// TIA Portal project "UsineEcole_TIAV20" (V20)

(* hardware
DEVICE "Station S71500/ET200MP_1"  S7-1500 station
   slot 0: "Châssis_0"  Rack  6ES7 590-1***0-0AA0
   slot 1: "PLC_1"  CPU 1518-4 PN/DP  6ES7 518-4AP00-0AB0  V2.9
      slot 3: "Ecran CPU_1"  6ES7591-1BA00-0AA0
      slot 32768: "Interface PROFINET_1"  X1
      slot 33024: "Interface PROFINET_2"  X2
      slot 33280: "Interface PROFINET GBIT_3"  X3
      slot 34817: "Virtual CP interface port_1"  Virtual CP interface port  Virtual CP interface port
   slot 2: "DI 32x24VDC HF_1"  DI 32x24VDC HF  6ES7 521-1BL00-0AB0  V2.1
   slot 3: "DQ 32x24VDC/0.5A ST_1"  DQ 32x24VDC/0.5A ST  6ES7 522-1BL00-0AB0  V2.0
DEVICE "Appareil GSD_1"  GSD.Device.PN
   slot 0: "Châssis"  Rack  V1.0
   slot 0: "REP 1"  AL1306  AL1306
      slot 0: "PROFINET interface"  PROFINET interface
      slot 1: "PN-IO"  PN-IO
         slot 1: "X21"  X21
         slot 2: "X22"  X22
   slot 1: "IO-Link  1 I Byte without PQI"  IO-Link  1 I Byte without PQI
   slot 1: "Digital Input"  Digital Input
   slot 1: "8 Ports - IO Mode_1"  8 Ports - IO Mode
      slot 0: "IO-Link Master Proxy"  IO-Link Master Proxy
   slot 1: "Digital Input without PD"  Digital Input without PD
   slot 2: "IO-Link  1 I Byte without PQI_1"  IO-Link  1 I Byte without PQI
   slot 2: "Digital Input_1"  Digital Input
   slot 2: "Digital Input without PD_1"  Digital Input without PD
   slot 3: "IO-Link  1 I Byte without PQI_2"  IO-Link  1 I Byte without PQI
   slot 3: "Digital Input_2"  Digital Input
   slot 3: "Digital Input without PD_2"  Digital Input without PD
   slot 4: "IO-Link  1 I Byte without PQI_3"  IO-Link  1 I Byte without PQI
   slot 4: "Digital Input_3"  Digital Input
   slot 4: "Digital Input without PD_3"  Digital Input without PD
   slot 5: "IO-Link  1 I Byte without PQI_4"  IO-Link  1 I Byte without PQI
   slot 5: "Digital Input_4"  Digital Input
   slot 5: "Digital Input without PD_4"  Digital Input without PD
   slot 6: "IO-Link  1 I Byte without PQI_5"  IO-Link  1 I Byte without PQI
   slot 6: "Digital Input_5"  Digital Input
   slot 6: "Digital Input without PD_5"  Digital Input without PD
   slot 7: "IO-Link  1 I Byte without PQI_6"  IO-Link  1 I Byte without PQI
   slot 7: "Digital Input_6"  Digital Input
   slot 7: "Digital Input without PD_6"  Digital Input without PD
   slot 8: "IO-Link  1 I Byte without PQI_7"  IO-Link  1 I Byte without PQI
   slot 8: "Digital Input_7"  Digital Input
   slot 8: "Digital Input without PD_7"  Digital Input without PD
DEVICE "Appareil GSD_2"  GSD.Device.PN
   slot 0: "Châssis"  Rack  V1.0
   slot 0: "REP 2"  AL1306  AL1306
      slot 0: "PROFINET interface"  PROFINET interface
      slot 1: "PN-IO"  PN-IO
         slot 1: "X21"  X21
         slot 2: "X22"  X22
   slot 1: "8 Ports - IO Mode_1"  8 Ports - IO Mode
      slot 0: "IO-Link Master Proxy"  IO-Link Master Proxy
   slot 1: "Digital Input without PD"  Digital Input without PD
   slot 2: "Digital Input without PD_1"  Digital Input without PD
   slot 3: "Digital Input without PD_2"  Digital Input without PD
   slot 4: "Digital Input without PD_3"  Digital Input without PD
   slot 5: "Digital Input without PD_4"  Digital Input without PD
   slot 6: "Digital Input without PD_5"  Digital Input without PD
   slot 7: "Digital Input without PD_6"  Digital Input without PD
   slot 8: "Digital Input without PD_7"  Digital Input without PD
DEVICE "Appareil GSD_3"  GSD.Device.PN
   slot 0: "Châssis"  Rack  V1.0
   slot 0: "REP 3"  AL1306  AL1306
      slot 0: "PROFINET interface"  PROFINET interface
      slot 1: "PN-IO"  PN-IO
         slot 1: "X21"  X21
         slot 2: "X22"  X22
   slot 1: "8 Ports - IO Mode_1"  8 Ports - IO Mode
      slot 0: "IO-Link Master Proxy"  IO-Link Master Proxy
   slot 1: "Digital Input without PD"  Digital Input without PD
   slot 2: "Digital Input without PD_1"  Digital Input without PD
   slot 3: "Digital Input without PD_2"  Digital Input without PD
   slot 4: "Digital Input without PD_3"  Digital Input without PD
   slot 5: "Digital Input without PD_4"  Digital Input without PD
   slot 6: "Digital Input without PD_5"  Digital Input without PD
   slot 7: "Digital Input without PD_6"  Digital Input without PD
   slot 8: "Digital Input without PD_7"  Digital Input without PD
DEVICE "Appareil GSD_4"  GSD.Device.PN
   slot 0: "Châssis"  Rack  V1.0
   slot 0: "REP 4"  AL1306  AL1306
      slot 0: "PROFINET interface"  PROFINET interface
      slot 1: "PN-IO"  PN-IO
         slot 1: "X21"  X21
         slot 2: "X22"  X22
   slot 1: "8 Ports - IO Mode_1"  8 Ports - IO Mode
      slot 0: "IO-Link Master Proxy"  IO-Link Master Proxy
   slot 1: "Digital Input without PD"  Digital Input without PD
   slot 2: "Digital Input without PD_1"  Digital Input without PD
   slot 3: "Digital Input without PD_2"  Digital Input without PD
   slot 4: "Digital Input without PD_3"  Digital Input without PD
   slot 5: "Digital Input without PD_4"  Digital Input without PD
   slot 6: "Digital Input without PD_5"  Digital Input without PD
   slot 7: "Digital Input without PD_6"  Digital Input without PD
   slot 8: "Digital Input without PD_7"  Digital Input without PD
DEVICE "Appareil GSD_5"  GSD.Device.PN
   slot 0: "Châssis"  Rack  V1.0
   slot 0: "REP 5"  AL1306  AL1306
      slot 0: "PROFINET interface"  PROFINET interface
      slot 1: "PN-IO"  PN-IO
         slot 1: "X21"  X21
         slot 2: "X22"  X22
   slot 1: "8 Ports - IO Mode_1"  8 Ports - IO Mode
      slot 0: "IO-Link Master Proxy"  IO-Link Master Proxy
   slot 1: "Digital Input without PD"  Digital Input without PD
   slot 2: "Digital Input without PD_1"  Digital Input without PD
   slot 3: "Digital Input without PD_2"  Digital Input without PD
   slot 4: "Digital Input without PD_3"  Digital Input without PD
   slot 5: "Digital Input without PD_4"  Digital Input without PD
   slot 6: "Digital Input without PD_5"  Digital Input without PD
   slot 7: "Digital Input without PD_6"  Digital Input without PD
   slot 8: "Digital Input without PD_7"  Digital Input without PD
DEVICE "Appareil GSD_6"  GSD.Device.PN
   slot 0: "Châssis"  Rack  V1.0
   slot 0: "REP 6"  AL1306  AL1306
      slot 0: "PROFINET interface"  PROFINET interface
      slot 1: "PN-IO"  PN-IO
         slot 1: "X21"  X21
         slot 2: "X22"  X22
   slot 1: "8 Ports - IO Mode_1"  8 Ports - IO Mode
      slot 0: "IO-Link Master Proxy"  IO-Link Master Proxy
   slot 1: "Digital Input without PD"  Digital Input without PD
   slot 2: "Digital Input without PD_1"  Digital Input without PD
   slot 3: "Digital Input without PD_2"  Digital Input without PD
   slot 4: "Digital Input without PD_3"  Digital Input without PD
   slot 5: "Digital Input without PD_4"  Digital Input without PD
   slot 6: "Digital Input without PD_5"  Digital Input without PD
   slot 7: "Digital Input without PD_6"  Digital Input without PD
   slot 8: "Digital Input without PD_7"  Digital Input without PD
DEVICE "Appareil GSD_7"  GSD.Device.PN
   slot 0: "Châssis"  Rack  V1.0
   slot 0: "Ilot 01"  EX260 SPN 1/2  EX260-SPN
      slot 0: "EX260 SPN 1/2"  EX260 SPN 1/2
      slot 1: "Interface"  Interface
         slot 1: "Port 1 - RJ45"  Port 1 - RJ45
         slot 2: "Port 2 - RJ45"  Port 2 - RJ45
      slot 1: "  4 byte  Output_1"    4 byte  Output
         slot 0: "  4 byte  Output"    4 byte  Output
DEVICE "Appareil GSD_8"  GSD.Device.PN
   slot 0: "Châssis"  Rack  V1.0
   slot 0: "ilot02"  EX260 SPN 1/2  EX260-SPN
      slot 0: "EX260 SPN 1/2"  EX260 SPN 1/2
      slot 1: "Interface"  Interface
         slot 1: "Port 1 - RJ45"  Port 1 - RJ45
         slot 2: "Port 2 - RJ45"  Port 2 - RJ45
      slot 1: "  4 byte  Output_1"    4 byte  Output
         slot 0: "  4 byte  Output"    4 byte  Output
DEVICE "Appareil GSD_9"  GSD.Device.PN
   slot 0: "Châssis"  Rack  V1.0
   slot 0: "SP-COP2-ENI"  R1.190.1320.0  R1.190.1320.0
      slot 0: "R1.190.1320.0"  R1.190.1320.0
      slot 1: "SP-COP2-ENI Diagnostics"  SP-COP2-ENI Diagnostics
      slot 2: "jz"  Interface
         slot 1: "RJ45 10/100 MBit/s"  RJ45 10/100 MBit/s
   slot 16: "Logic input block 1_1"  Logic input block 1
      slot 0: "Logic input block 1"  Logic input block 1
   slot 21: "Logic output block 1_1"  Logic output block 1
      slot 0: "Logic output block 1"  Logic output block 1
   slot 32: "CRC data_1"  CRC data
      slot 0: "CRC data"  CRC data
   slot 33: "Status data_1"  Status data
      slot 0: "Status data"  Status data
   slot 34: "Auxiliary data_1"  Auxiliary data
      slot 0: "Auxiliary data"  Auxiliary data
DEVICE "HMI_1"  TP1500 Comfort
   slot 0: "HMI_1"  TP1500 Comfort  6AV2 124-0QC02-0AX1  17.0.0.0
   slot 1: "HMI_RT_1"  TP1500 Comfort  6AV2 124-0QC02-0AX1  17.0.0.0
   slot 5: "HMI_1.IE_CP_1"  PROFINET Interface  17.0.0.0
      slot 1: "Interface PROFINET_1"  PROFINET Interface
         slot 1: "Port_1"  Port
         slot 2: "Port_2"  Port
   slot 6: "HMI_1.IE_CP_2"  PROFINET Interface  17.0.0.0
      slot 1: "Interface PROFINET_GBit"  PROFINET Interface
         slot 1: "Port_1"  Port
   slot 7: "HMI_1.MPI/DP_CP_1"  MPI/DP Interface  17.0.0.0
DEVICE "SINAMICS G_1"  Sinamics.Device
   slot 0: "	_0"  Rail  SinamicsG120CRackP
   slot 0: "Convoyeur 01"  G120C PN  6SL3210-1KE11-8UF2  4.7.13
      slot 1: "Interface PROFINET"  MDD-SinamicsG120-P
      slot 3: "PM G120C"  PM G120C  6SL3210-1KE11-8UF2  -
DEVICE "SINAMICS G_2"  Sinamics.Device
   slot 0: "	_0"  Rail  SinamicsG120CRackP
   slot 0: "Convoyeur 02"  G120C PN  6SL3210-1KE11-8UF2  4.7.13
      slot 1: "Interface PROFINET"  MDD-SinamicsG120-P
      slot 3: "PM G120C"  PM G120C  6SL3210-1KE11-8UF2  -
DEVICE "SINAMICS G_3"  Sinamics.Device
   slot 0: "	_0"  Rail  SinamicsG120CRackP
   slot 0: "Convoyeur 03"  G120C PN  6SL3210-1KE11-8UF2  4.7.13
      slot 1: "Interface PROFINET"  MDD-SinamicsG120-P
      slot 3: "PM G120C"  PM G120C  6SL3210-1KE11-8UF2  -
DEVICE "Appareil GSD_10"  GSD.Device
   slot 0: "Châssis_0"  Rail
DEVICE "Appareil GSD_12"  GSD.Device.PN
   slot 0: "Châssis"  Rack  V1.0
   slot 0: "UR_R4"  V1.0  0000201
      slot 0: "V1.0"  V1.0
      slot 1: "Interface"  Interface
         slot 1: "RJ45 10/100 MBit/s"  RJ45 10/100 MBit/s
   slot 1: "1_T2O State_1"  1_T2O State  1.0
      slot 0: "1_T2O State"  1_T2O State
   slot 2: "2_T2O IO_1"  2_T2O IO  1.0
      slot 0: "2_T2O IO"  2_T2O IO
   slot 3: "3_T2O Joints_1"  3_T2O Joints  1.0
      slot 0: "3_T2O Joints"  3_T2O Joints
   slot 4: "4_T2O TCP_1"  4_T2O TCP  1.0
      slot 0: "4_T2O TCP"  4_T2O TCP
   slot 5: "5_T2O General Purpose Bit Registers_1"  5_T2O General Purpose Bit Registers  1.0
      slot 0: "5_T2O General Purpose Bit Registers"  5_T2O General Purpose Bit Registers
   slot 6: "6_T2O General Purpose Int Registers_1"  6_T2O General Purpose Int Registers  1.0
      slot 0: "6_T2O General Purpose Int Registers"  6_T2O General Purpose Int Registers
   slot 7: "7_T2O General Purpose Float Registers_1"  7_T2O General Purpose Float Registers  1.0
      slot 0: "7_T2O General Purpose Float Registers"  7_T2O General Purpose Float Registers
   slot 8: "8_O2T Robot IO_1"  8_O2T Robot IO  1.0
      slot 0: "8_O2T Robot IO"  8_O2T Robot IO
   slot 9: "9_O2T General Purpose Registers 1_1"  9_O2T General Purpose Registers 1  1.0
      slot 0: "9_O2T General Purpose Registers 1"  9_O2T General Purpose Registers 1
   slot 10: "10_O2T General Purpose Registers 2_1"  10_O2T General Purpose Registers 2  1.0
      slot 0: "10_O2T General Purpose Registers 2"  10_O2T General Purpose Registers 2
DEVICE "Appareil GSD_13"  GSD.Device.PN
   slot 0: "Châssis"  Rack  V1.0
   slot 0: "URIODev1_1"  V1.0  0000201
      slot 0: "V1.0"  V1.0
      slot 1: "Interface"  Interface
         slot 1: "RJ45 10/100 MBit/s"  RJ45 10/100 MBit/s
   slot 1: "1_T2O State_1"  1_T2O State  1.0
      slot 0: "1_T2O State"  1_T2O State
   slot 2: "2_T2O IO_1"  2_T2O IO  1.0
      slot 0: "2_T2O IO"  2_T2O IO
   slot 3: "3_T2O Joints_1"  3_T2O Joints  1.0
      slot 0: "3_T2O Joints"  3_T2O Joints
   slot 4: "4_T2O TCP_1"  4_T2O TCP  1.0
      slot 0: "4_T2O TCP"  4_T2O TCP
   slot 5: "5_T2O General Purpose Bit Registers_1"  5_T2O General Purpose Bit Registers  1.0
      slot 0: "5_T2O General Purpose Bit Registers"  5_T2O General Purpose Bit Registers
   slot 6: "6_T2O General Purpose Int Registers_1"  6_T2O General Purpose Int Registers  1.0
      slot 0: "6_T2O General Purpose Int Registers"  6_T2O General Purpose Int Registers
   slot 7: "7_T2O General Purpose Float Registers_1"  7_T2O General Purpose Float Registers  1.0
      slot 0: "7_T2O General Purpose Float Registers"  7_T2O General Purpose Float Registers
   slot 8: "8_O2T Robot IO_1"  8_O2T Robot IO  1.0
      slot 0: "8_O2T Robot IO"  8_O2T Robot IO
   slot 9: "9_O2T General Purpose Registers 1_1"  9_O2T General Purpose Registers 1  1.0
      slot 0: "9_O2T General Purpose Registers 1"  9_O2T General Purpose Registers 1
   slot 10: "10_O2T General Purpose Registers 2_1"  10_O2T General Purpose Registers 2  1.0
      slot 0: "10_O2T General Purpose Registers 2"  10_O2T General Purpose Registers 2
   slot 11: "PROFIsafe_1"  PROFIsafe  1.0
      slot 0: "Module Access Point"  Module Access Point
DEVICE "Appareil GSD_11"  GSD.Device.PN
   slot 0: "Châssis"  Rack  V1.0
   slot 0: "CP-1604"  V2.5  A05B-2500-J930  V2.5
      slot 0: "CP 1604"  CP 1604
      slot 1: "Interface"  Interface
         slot 1: "Port_1"  Port
   slot 1: "  32 octets_1"  32 bytes  1.0
      slot 0: "  32 octets"  32 bytes
DEVICE "Appareil GSD_14"  GSD.Device.PN
   slot 0: "Châssis"  Rack  V1.0
   slot 0: "cv-x400"  CV-X4XX  CV-X4XX  5.1
      slot 0: "CV-X4XX"  CV-X4XX  5.1
      slot 1: "Interface"  Interface
         slot 1: "Port 1"  Port 1
   slot 1: "Command and Result Status_1"  Command and Result Status
      slot 0: "Command and Result Status"  Command and Result Status
   slot 2: "Trg Ready Status_1"  Trg Ready Status
      slot 0: "Trg Ready Status"  Trg Ready Status
   slot 3: "Trg Ack Status_1"  Trg Ack Status
      slot 0: "Trg Ack Status"  Trg Ack Status
   slot 4: "Miscellaneous Status_1"  Miscellaneous Status
      slot 0: "Miscellaneous Status"  Miscellaneous Status
   slot 5: "Tool Judge Value_1"  Tool Judge Value
      slot 0: "Tool Judge Value"  Tool Judge Value
   slot 6: "Result Data 128Byte_1"  Result Data 128Byte
      slot 0: "Result Data 128Byte"  Result Data 128Byte
   slot 7: "Result Data 32Byte_1"  Result Data 32Byte
      slot 0: "Result Data 32Byte"  Result Data 32Byte
   slot 8: "Result Data 32Byte_2"  Result Data 32Byte
      slot 0: "Result Data 32Byte"  Result Data 32Byte
   slot 9: "Result Data 32Byte_3"  Result Data 32Byte
      slot 0: "Result Data 32Byte"  Result Data 32Byte
   slot 10: "Result Data 32Byte_4"  Result Data 32Byte
      slot 0: "Result Data 32Byte"  Result Data 32Byte
   slot 11: "Result Data 32Byte_5"  Result Data 32Byte
      slot 0: "Result Data 32Byte"  Result Data 32Byte
   slot 12: "Command and Result Control_1"  Command and Result Control
      slot 0: "Command and Result Control"  Command and Result Control
   slot 13: "Trg Control_1"  Trg Control
      slot 0: "Trg Control"  Trg Control
   slot 14: "Miscellaneous Control_1"  Miscellaneous Control
      slot 0: "Miscellaneous Control"  Miscellaneous Control
   slot 15: "Reserved Control_1"  Reserved Control
      slot 0: "Reserved Control"  Reserved Control
   slot 16: "Reserved Control_2"  Reserved Control
      slot 0: "Reserved Control"  Reserved Control
   slot 17: "Parameter 128Byte_1"  Parameter 128Byte
      slot 0: "Parameter 128Byte"  Parameter 128Byte
   slot 18: "Parameter 32Byte_1"  Parameter 32Byte
      slot 0: "Parameter 32Byte"  Parameter 32Byte
   slot 19: "Parameter 32Byte_2"  Parameter 32Byte
      slot 0: "Parameter 32Byte"  Parameter 32Byte
   slot 20: "Parameter 32Byte_3"  Parameter 32Byte
      slot 0: "Parameter 32Byte"  Parameter 32Byte
   slot 21: "Parameter 32Byte_4"  Parameter 32Byte
      slot 0: "Parameter 32Byte"  Parameter 32Byte
   slot 22: "Parameter 32Byte_5"  Parameter 32Byte
      slot 0: "Parameter 32Byte"  Parameter 32Byte
DEVICE "GSD device_1"  GSD.Device.PN
   slot 0: "Rack"  Rack  V1.0
   slot 0: "REP 4_rep"  AL1102  AL1102
      slot 0: "AL1102"  AL1102
      slot 1: "X1"  X1
         slot 1: "Port 1"  Port 1
         slot 2: "Port 2"  Port 2
      slot 1: "8 Ports_1"  8 Ports  AL1102
         slot 0: "IO-Link Master"  IO-Link Master
   slot 1: "Digital Input + PQI"  Digital Input + PQI
   slot 2: "Digital Input + PQI_1"  Digital Input + PQI
DEVICE "GSD device_2"  GSD.Device.PN
   slot 0: "Rack"  Rack  V1.0
   slot 0: "OmniCore"  OmniCore Standard  3020-x  V1.1
      slot 0: "OmniCore Standard PROFINET Device"  OmniCore Standard PROFINET Device
      slot 1: "PROFINET Interface"  PROFINET Interface
         slot 1: "Network Port 1"  Network Port 1
   slot 1: "DI 8 bytes_1"  DI 8 bytes
      slot 0: "DI 8 bytes"  DI 8 bytes
   slot 2: "DO 8 bytes_1"  DO 8 bytes
      slot 0: "DO 8 bytes"  DO 8 bytes
*)

// ===== PLC "PLC_1"  CPU 1518-4 PN/DP =====

VAR_GLOBAL   // PLC tag table "Table de variables standard"
   "I_En_Service" AT %I0.0 : Bool;
   "I_Not_AU" AT %I0.1 : Bool;   // Entree AU: 1 = pas d'arret d'urgence
   "I_En_Manuel" AT %I0.2 : Bool;
   "I_En_Automatique" AT %I0.3 : Bool;
   "I_porte_non_réarmée" AT %I0.4 : Bool;
   "I_porte_01_Op" AT %I0.5 : Bool;
   "I_porte_02_Op" AT %I0.6 : Bool;
   "I_libre_I07" AT %I0.7 : Bool;
   "I_libre_I10" AT %I1.0 : Bool;
   "I_Def_Thermique_CV01_hyppo" AT %I1.1 : Bool;
   "I_Def_Thermique_CV02_hyppo" AT %I1.2 : Bool;
   "I_Def_Thermique_CV03_hyppo" AT %I1.3 : Bool;
   "I_Def_Thermique_CV04_hyppo" AT %I1.4 : Bool;
   "I_libre_I15" AT %I1.5 : Bool;
   "I_libre_I16" AT %I1.6 : Bool;
   "I_libre_I17" AT %I1.7 : Bool;
   "I_libre_I20" AT %I2.0 : Bool;
   "I_libre_I21" AT %I2.1 : Bool;
   "I_libre_I22" AT %I2.2 : Bool;
   "I_libre_I23" AT %I2.3 : Bool;
   "I_libre_I24" AT %I2.4 : Bool;
   "I_libre_I25" AT %I2.5 : Bool;
   "I_libre_I26" AT %I2.6 : Bool;
   "I_libre_I27" AT %I2.7 : Bool;
   "I_libre_I30" AT %I3.0 : Bool;
   "I_libre_I31" AT %I3.1 : Bool;
   "I_libre_I32" AT %I3.2 : Bool;
   "I_libre_I33" AT %I3.3 : Bool;
   "I_libre_I34" AT %I3.4 : Bool;
   "I_libre_I35" AT %I3.5 : Bool;
   "I_libre_I36" AT %I3.6 : Bool;
   "I_libre_I37" AT %I3.7 : Bool;
   "I_Pres_Pal_B01" AT %I5.0 : Bool;
   "I_Pres_Elev_B01" AT %I4.0 : Bool;
   "I_Elev_01_Bas" AT %I5.1 : Bool;
   "I_Elev_01_Haut" AT %I4.1 : Bool;
   "I_Pres_Pal_B02" AT %I5.2 : Bool;
   "I_Pres_Elev_B02" AT %I4.2 : Bool;
   "I_Elev_02_Bas" AT %I5.3 : Bool;
   "I_Elev_02_Haut" AT %I4.3 : Bool;
   "I_Pres_Pal_B03" AT %I5.4 : Bool;
   "I_Pres_Elev_B03" AT %I4.4 : Bool;
   "I_Elev_03_Bas" AT %I5.5 : Bool;
   "I_Elev_03_Haut" AT %I4.5 : Bool;
   "I_Pres_Pal_B04" AT %I5.6 : Bool;
   "I_Pres_Elev_B04" AT %I4.6 : Bool;
   "I_Elev_04_Bas" AT %I5.7 : Bool;
   "I_Elev_04_Haut" AT %I4.7 : Bool;
   "I_Pres_Pal_B05" AT %I7.0 : Bool;
   "I_Pres_Elev_B05" AT %I6.0 : Bool;
   "I_Elev_05_Bas" AT %I7.1 : Bool;
   "I_Elev_05_Haut" AT %I6.1 : Bool;
   "I_Pres_Pal_B06" AT %I7.2 : Bool;
   "I_Pres_Elev_B06" AT %I6.2 : Bool;
   "I_Elev_06_Bas" AT %I7.3 : Bool;
   "I_Elev_06_Haut" AT %I6.3 : Bool;
   "I_Pres_Pal_B07" AT %I7.4 : Bool;
   "I_Pres_Elev_B07" AT %I6.4 : Bool;
   "I_Elev_07_Bas" AT %I7.5 : Bool;
   "I_Elev_07_Haut" AT %I6.5 : Bool;
   "I_det_Phot_01" AT %I11.0 : Bool;
   "I_det_Phot_02" AT %I10.0 : Bool;
   "I_det_Phot_03" AT %I11.1 : Bool;
   "I_verin_blocage_boite_sorti_01" AT %I10.1 : Bool;
   "I_verin_blocage_boite_rentré_01" AT %I11.2 : Bool;
   "I_verin_blocage_boite_sorti_02" AT %I10.2 : Bool;
   "I_verin_blocage_boite_sorti_03" AT %I10.3 : Bool;
   "I_verin_blocage_boite_rentré_03" AT %I11.4 : Bool;
   "I_verin_blocage_boite_rentré_02" AT %I11.3 : Bool;
   "I_verin_blocage_boite_sorti_04" AT %I10.4 : Bool;
   "I_verin_blocage_boite_rentré_04" AT %I11.5 : Bool;
   "I_Det_Phot_04" AT %I13.0 : Bool;
   "I_Det_Phot_05" AT %I12.0 : Bool;
   "I_Det_Phot_06" AT %I13.1 : Bool;
   "I_Det_Photo_7" AT %I15.0 : Bool;
   "I_Det_Photo_8" AT %I14.0 : Bool;
   "I_Det_Photo_9" AT %I15.1 : Bool;
   "I_Wieland_Au_armoire" AT %I16.0 : Bool;
   "I_Wieland_Au_porte01" AT %I16.1 : Bool;
   "I_Wieland_Au_Porte02" AT %I16.2 : Bool;
   "I_Wieland_Au_Robot01_Fanuc" AT %I16.3 : Bool;
   "I_Wieland_Au_Robot02_Fanuc" AT %I16.4 : Bool;
   "I_Wieland_Au_Robot03_ABB" AT %I16.5 : Bool;
   "I_Wielmand_Au_Robot04_UR" AT %I16.6 : Bool;
   "I_Wieland_Au_Robot05_UR" AT %I16.7 : Bool;
   "I_wieland_Au_Carroussel" AT %I17.0 : Bool;
   "I_Wieland_Au_Carterisation" AT %I17.1 : Bool;
   "I_Wieland_Porte 01 ouverte" AT %I17.2 : Bool;
   "I_Wieland_Porte 02 Ouverte" AT %I17.3 : Bool;
   "I_Wieland_Rearmement" AT %I17.4 : Bool;
   "I_Wieland_Dmd acces" AT %I17.5 : Bool;
   "I_Wieland_Mise sous puissance" AT %I17.6 : Bool;
   "I_Wieland_Mise hors puissance" AT %I17.7 : Bool;
   "I_Wieland_Acces_autorisé" AT %I18.0 : Bool;
   "I_Wieland_rearmement_Porte" AT %I18.1 : Bool;
   "I_Wieland_En_Service" AT %I18.2 : Bool;
   "I_Wieland_Porte_non_Réarmée" AT %I18.3 : Bool;
   "I_porte_vision_op" AT %I7.6 : Bool;
   "I_porte_vision_cl" AT %I6.6 : Bool;
   "Tag_1" AT %I590.0 : Bool;
   "Tag_2" AT %I590.1 : Bool;
   "UR01I" AT %I556.0 : "UR__T2O_IOs";
   "Fanuc01_Selecteur_Auto" AT %I30.4 : Bool;
   "Fanuc02_Selecteur_Auto" AT %I220.4 : Bool;
   "Fanuc02_reception_signal_pret" AT %I30.5 : Bool;
   "Fanuc01_reception_signal_pret" AT %I220.5 : Bool;
   "VisionOK" AT %I42.0 : Bool;   // vision OK
   "Tag_8" AT %I42.1 : Bool;
   "Tag_9" AT %I42.2 : Bool;
   "Tag_10" AT %I7.7 : Bool;
   "O_CL_verte" AT %Q0.0 : Bool;
   "O_CL_Orange" AT %Q0.1 : Bool;
   "O_CL_Rouge" AT %Q0.2 : Bool;
   "Q_LibreQ03" AT %Q0.3 : Bool;
   "Q_LibreQ04" AT %Q0.4 : Bool;
   "Q_LibreQ05" AT %Q0.5 : Bool;
   "Q_LibreQ06" AT %Q0.6 : Bool;
   "Q_LibreQ07" AT %Q0.7 : Bool;
   "Q_LibreQ10" AT %Q1.0 : Bool;
   "Q_LibreQ11" AT %Q1.1 : Bool;
   "Q_LibreQ12" AT %Q1.2 : Bool;
   "Q_LibreQ13" AT %Q1.3 : Bool;
   "Q_LibreQ14" AT %Q1.4 : Bool;
   "Q_LibreQ15" AT %Q1.5 : Bool;
   "Q_LibreQ16" AT %Q1.6 : Bool;
   "Q_LibreQ17" AT %Q1.7 : Bool;
   "O_ON_CV_01_Hyppo" AT %Q2.0 : Bool;
   "O_ON_CV_02_Hyppo" AT %Q2.1 : Bool;
   "O_ON_CV_03_Hyppo" AT %Q2.2 : Bool;
   "O_ON_CV_04_Hyppo" AT %Q2.3 : Bool;
   "Q_LibreQ24" AT %Q2.4 : Bool;
   "Q_LibreQ25" AT %Q2.5 : Bool;
   "Q_LibreQ26" AT %Q2.6 : Bool;
   "Q_LibreQ27" AT %Q2.7 : Bool;
   "Q_LibreQ30" AT %Q3.0 : Bool;
   "Q_LibreQ31" AT %Q3.1 : Bool;
   "Q_LibreQ32" AT %Q3.2 : Bool;
   "Q_LibreQ33" AT %Q3.3 : Bool;
   "Q_LibreQ34" AT %Q3.4 : Bool;
   "Q_LibreQ35" AT %Q3.5 : Bool;
   "Q_LibreQ36" AT %Q3.6 : Bool;
   "Q_LibreQ37" AT %Q3.7 : Bool;
   "O_Rentrer_Butée_01" AT %Q10.0 : Bool;
   "O_Rentrer_Butée_EL_01" AT %Q10.1 : Bool;
   "O_Monter_EL_01" AT %Q10.2 : Bool;
   "O_Desc_EL_01" AT %Q10.3 : Bool;
   "O_Rentrer_Butée_02" AT %Q10.4 : Bool;
   "O_Rentrer_Butée_EL_02" AT %Q10.5 : Bool;
   "O_Monter_EL_02" AT %Q10.6 : Bool;
   "O_Desc_EL_02" AT %Q10.7 : Bool;
   "O_Rentrer_Butée_03" AT %Q11.0 : Bool;
   "O_Rentrer_Butée_EL_03" AT %Q11.1 : Bool;
   "O_Monter_EL_03" AT %Q11.2 : Bool;
   "O_Desc_EL_03" AT %Q11.3 : Bool;
   "O_Rentrer_Butée_04" AT %Q11.4 : Bool;
   "O_Rentrer_Butée_EL_04" AT %Q11.5 : Bool;
   "O_Monter_EL_04" AT %Q11.6 : Bool;
   "O_Desc_EL_04" AT %Q11.7 : Bool;
   "O_Rentrer_Butée_05" AT %Q12.0 : Bool;
   "O_Rentrer_Butée_EL_05" AT %Q12.1 : Bool;
   "O_Monter_EL_05" AT %Q12.2 : Bool;
   "O_Desc_EL_05" AT %Q12.3 : Bool;
   "O_Rentrer_Butée_06" AT %Q12.4 : Bool;
   "O_Rentrer_Butée_EL_06" AT %Q12.5 : Bool;
   "O_Monter_EL_06" AT %Q12.6 : Bool;
   "O_Desc_EL_06" AT %Q12.7 : Bool;
   "O_Rentrer_Butée_07" AT %Q13.0 : Bool;
   "O_Rentrer_Butée_EL_07" AT %Q13.1 : Bool;
   "O_Monter_EL_07" AT %Q13.2 : Bool;
   "O_Desc_EL_07" AT %Q13.3 : Bool;
   "O_Sortir_Blocage_boite_01" AT %Q14.0 : Bool;
   "O_Rentrer_Blocage_boite_01" AT %Q14.1 : Bool;
   "O_Sortir_Blocage_boite_02" AT %Q14.2 : Bool;
   "O_Sortir_Blocage_boite_03" AT %Q14.4 : Bool;
   "O_Sortir_Blocage_boite_04" AT %Q14.6 : Bool;
   "O_Rentrer_Blocage_boite_02" AT %Q14.3 : Bool;
   "O_Rentrer_Blocage_boite_03" AT %Q14.5 : Bool;
   "O_Rentrer_Blocage_boite_04" AT %Q14.7 : Bool;
   "O_Op_Porte_Vision" AT %Q13.4 : Bool;
   "O_Cl_porte_Vision" AT %Q13.5 : Bool;
   "Q_Wieland_Acces_Autorisé" AT %Q18.0 : Bool;
   "O_trigger_CVX" AT %Q69.0 : Bool;
   "UR01O" AT %Q396.0 : "UR__O2T_IOs";
   "Tag_3" AT %Q420.0 : Bool;
   "Tag_4" AT %Q420.1 : Bool;
   "Tag_5" AT %Q420.2 : Bool;
   "Tag_6" AT %Q644.2 : Bool;
   "Fanuc01_Autor_Prise" AT %Q40.5 : Bool;
   "Fanuc02_Autor_Prise" AT %Q31.5 : Bool;
   "Fanuc02_Autor_Depose" AT %Q31.6 : Bool;
   "Fanuc01_envoi_signal_pret_vers_fanuc02" AT %Q31.7 : Bool;
   "Fanuc02_envoi_signal_pret_vers_fanuc_01" AT %Q40.6 : Bool;
   "Defaut_EL01" AT %M20.0 : Bool;
   "Defaut_EL02" AT %M20.1 : Bool;
   "Defaut_EL03" AT %M20.2 : Bool;
   "Defaut_EL04" AT %M20.3 : Bool;
   "Defaut_EL05" AT %M20.4 : Bool;
   "Defaut_EL06" AT %M20.5 : Bool;
   "Defaut_EL07" AT %M20.6 : Bool;
   "System_Byte" AT %MB1 : Byte;
   "FirstScan" AT %M1.0 : Bool;
   "DiagStatusUpdate" AT %M1.1 : Bool;
   "AlwaysTRUE" AT %M1.2 : Bool;
   "AlwaysFALSE" AT %M1.3 : Bool;
   "Clock_Byte" AT %MB0 : Byte;
   "Clock_10Hz" AT %M0.0 : Bool;
   "Clock_5Hz" AT %M0.1 : Bool;
   "Clock_2.5Hz" AT %M0.2 : Bool;
   "Clock_2Hz" AT %M0.3 : Bool;
   "Clock_1.25Hz" AT %M0.4 : Bool;
   "Clock_1Hz" AT %M0.5 : Bool;
   "Clock_0.625Hz" AT %M0.6 : Bool;
   "Clock_0.5Hz" AT %M0.7 : Bool;
   "O_On_CV01" AT %M30.0 : Bool;
   "O_On_CV02" AT %M30.1 : Bool;
   "O_On_CV03" AT %M30.2 : Bool;
   "B_autorisation_depose_CV02" AT %M40.0 : Bool;
   "B_autorisation_prise_CV02" AT %M40.1 : Bool;
   "Step_CV02" AT %MW50 : Int;
   "Step_CV03" AT %MW51 : Int;
   "B_autorisation_prise_CV03" AT %M40.2 : Bool;
   "B_autorisation_depose_CV03" AT %M40.3 : Bool;
   "O_On_CV01_TP_Robot" AT %M100.0 : Bool;
   "Fanuc01_Fanuc02_En_Auto" AT %M200.0 : Bool;
END_VAR

VAR_GLOBAL   // PLC tag table "UR_R4_tags"
   "UR1_Robot_status" AT %I556.0 : "UR_1_T2O_State";
   "UR1_IO_status" AT %I588.0 : "UR_2_T2O_IO";
   "UR1_Joints" AT %I656.0 : "UR_3_T2O_Joints";
   "UR1_TCP" AT %I760.0 : "UR_4_T2O_TCP";
   "UR1_Bit_registers" AT %I50.0 : "UR_5_T2O_BitRegisters";
   "UR1_Int_registers" AT %I836.0 : "UR_6_T2O_IntRegisters";
   "UR1_Float_registers" AT %I932.0 : "UR_7_T2O_FloatRegisters";
   "UR1_Robot_IO_Q" AT %Q396.0 : "UR_8_O2T_Robot_IO";
   "UR1_Registers_1_Q" AT %Q420.0 : "UR_9_O2T_Registers";
   "UR1_Registers_2_Q" AT %Q520.0 : "UR_9_O2T_Registers";
END_VAR

VAR_GLOBAL   // PLC tag table "UR_R5_tags"
   "UR2_Robot_status" AT %I1028.0 : "UR_1_T2O_State";
   "UR2_IO_status" AT %I1060.0 : "UR_2_T2O_IO";
   "UR2_Joints" AT %I1128.0 : "UR_3_T2O_Joints";
   "UR2_TCP" AT %I1232.0 : "UR_4_T2O_TCP";
   "UR2_Bit_registers" AT %I58.0 : "UR_5_T2O_BitRegisters";
   "UR2_Int_registers" AT %I1308.0 : "UR_6_T2O_IntRegisters";
   "UR2_Float_registers" AT %I1404.0 : "UR_7_T2O_FloatRegisters";
   "UR2_Robot_IO_Q" AT %Q620.0 : "UR_8_O2T_Robot_IO";
   "UR2_Registers_1_Q" AT %Q644.0 : "UR_9_O2T_Registers";
   "UR2_Registers_2_Q" AT %Q744.0 : "UR_9_O2T_Registers";
END_VAR

VAR_GLOBAL   // PLC tag table "FANUC_R1_tags"
   "I_FANUC_R1" AT %I218.0 : "Fanuc_status";
   "O_FANUC_R1_IMSTP" AT %Q36.0 : Bool;
   "O_FANUC_R1_Fault_reset" AT %Q36.1 : Bool;
   "O_FANUC_R1_Start_Pns_strobe" AT %Q36.2 : Bool;
   "O_FANUC_R1_Enable" AT %Q36.3 : Bool;
   "O_FANUC_R1_PNS1" AT %Q36.4 : Bool;
   "O_FANUC_R1_PNS2" AT %Q36.5 : Bool;
   "O_FANUC_R1_Cicle_stop" AT %Q36.6 : Bool;   // ABORT ALL
   "O_FANUC_R1_Autor_Prise" AT %Q36.7 : Bool;
   "O_FANUC_R1_Autor_Depose" AT %Q37.0 : Bool;
   "O_FANUC_R1_HOME" AT %Q37.1 : Bool;
   "O_FANUC_R1" AT %Q36.0 : "Fanuc_cmd";
END_VAR

VAR_GLOBAL   // PLC tag table "FANUC_R2_tags"
   "I_FANUC_R2_Cmd_enabled" AT %I28.0 : Bool;
   "I_FANUC_R2_FAULT" AT %I28.1 : Bool;
   "I_FANUC_R2_Prog_running" AT %I28.2 : Bool;
   "I_FANUC_R2_Snack" AT %I28.3 : Bool;
   "I_FANUC_R2_Teach_on" AT %I28.4 : Bool;
   "I_FANUC_R2_In_auto" AT %I28.5 : Bool;
   "I_FANUC_R2_Libre" AT %I28.6 : Bool;
   "I_FANUC_R2_Libre_1" AT %I28.7 : Bool;
   "I_FANUC_R2_Fin_prise" AT %I29.0 : Bool;
   "I_FANUC_R2_Fin_depose" AT %I29.1 : Bool;
   "I_FANUC_R2" AT %I28.0 : "Fanuc_status";
   "O_FANUC_R2_IMSTP" AT %Q28.0 : Bool;
   "O_FANUC_R2_Fault_reset" AT %Q28.1 : Bool;
   "O_FANUC_R2_Start_Pns_strobe" AT %Q28.2 : Bool;
   "O_FANUC_R2_Enable" AT %Q28.3 : Bool;
   "O_FANUC_R2_PNS1" AT %Q28.4 : Bool;
   "O_FANUC_R2_PNS2" AT %Q28.5 : Bool;
   "O_FANUC_R2_Cicle_stop" AT %Q28.6 : Bool;   // ABORT ALL
   "O_FANUC_R2_Autor_Prise" AT %Q28.7 : Bool;
   "O_FANUC_R2_Autor_Depose" AT %Q29.0 : Bool;
   "O_FANUC_R2_HOME" AT %Q29.1 : Bool;
   "O_FANUC_R2" AT %Q28.0 : "Fanuc_cmd";
END_VAR

VAR_GLOBAL   // PLC tag table "CV01_conditionnement"
   "CV01_Status" AT %I256.0 : "Var_G120C_status";
   "CV01_Cmd" AT %Q256.0 : "Var_G120C_cmd";
END_VAR

VAR_GLOBAL   // PLC tag table "CV02_conditionnement"
   "CV02_Status" AT %I260.0 : "Var_G120C_status";
   "CV02_Cmd" AT %Q260.0 : "Var_G120C_cmd";
END_VAR

VAR_GLOBAL   // PLC tag table "CV03_conditionnement"
   "CV03_Status" AT %I264.0 : "Var_G120C_status";
   "CV03_Cmd" AT %Q264.0 : "Var_G120C_cmd";
END_VAR

VAR_GLOBAL   // PLC tag table "GoFa_R3_tags"
   "I_GoFa" AT %I1500.0 : "GoFa_Status";
   "O_GoFa" AT %Q240.0 : "GoFa_cmd";
END_VAR

TYPE "Variateur_G120C"
VERSION : 0.1
   STRUCT
      Reserve01 : Bool;
      Reserve02 : Bool;
      PilotageParApi : Bool;
      InversionConsigne : Bool;
      Reserve03 : Bool;
      PotPlus : Bool;
      PotMoins : Bool;
      Reserve04 : Bool;
      Marche : Bool;
      Arret2 : Bool;
      Arret3 : Bool;
      DebloqFonctionnement : Bool;
      DebloqRampe : Bool;
      GelerGenerateurRampe : Bool;
      DebloqConsigne : Bool;
      AcquitDefaut : Bool;
      Consigne : Int;
      EcartVitesse : Bool;
      CommandeDemander : Bool;
      VitesseMaxAtteinte : Bool;
      Limite : Bool;
      FreinMoteur : Bool;
      AlarmeSurchauffe : Bool;
      MoteurSensAvant : Bool;
      SurchargeMoteur : Bool;
      PretEnclenchement : Bool;
      PretFonctionnement : Bool;
      Fonctionnement_Debloq : Bool;
      DefautActif : Bool;
      Arret2Etat : Bool;
      Arret3Etat : Bool;
      BlocageActif : Bool;
      AlarmeActive : Bool;
      Vitesse : Int;
   END_STRUCT;
END_TYPE

TYPE "Imprimante3D"
VERSION : 0.1
   STRUCT
      Status : Struct
         x_Ready : Bool;
         x_Busy : Bool;
         x_Work_done : Bool;
         x_Work_done_manu : Bool;
         x_AtHome : Bool;
         x_HasPrintSurface : Bool;
         t_Elapsed_time : Time;
         t_Remaining_time : Time;
         x_Fault : Time;
      END_STRUCT;
      Cmd : Struct
         x_Start : Bool;
         x_Stop : Bool;
         x_Resume : Bool;
         x_Home : Bool;
      END_STRUCT;
      Printer_ID : Int;
   END_STRUCT;
END_TYPE

TYPE "Convoyeur_Hipp"
VERSION : 0.1
   STRUCT
      Status : Struct
         x_EnMarche : Bool;
         x_Fault : Bool;
      END_STRUCT;
      Cmd : Struct
         x_Start : Bool;
         x_Stop : Bool;
      END_STRUCT;
   END_STRUCT;
END_TYPE

TYPE "Station_Hipp"
VERSION : 0.1
   STRUCT
      Elevateur : Struct
         status : Struct
            x_Pos_haute : Bool;
            x_Pos_basse : Bool;
            x_Pres_palette : Bool;
            x_Busy : Bool;
            x_Free : Bool;
            x_Await_work_done : Bool;
            x_Has_print_surface : Bool;
            x_Has_3D_piece : Bool;
            x_Piece_control_OK : Bool;
            x_Print_surface_clean : Bool;
            x_Fault : Bool;
         END_STRUCT;
         cmd : Struct
            x_Elevator_up : Bool;
            x_Elevator_down : Bool;
            x_Stopper_down : Bool;
            x_Elevator_up_manual : Bool;
            x_Elevator_down_manual : Bool;
            x_Stopper_down_manual : Bool;
         END_STRUCT;
      END_STRUCT;
      Buffer : Struct
         status : Struct
            x_Pres_palette : Bool;
            x_buffer_full : Bool;
            x_fault : Bool;
         END_STRUCT;
         cmd : Struct
            x_Stopper_down : Bool;
            x_Stopper_down_manu : Bool;
         END_STRUCT;
      END_STRUCT;
      Num_station : Int;
   END_STRUCT;
END_TYPE

TYPE "Fanuc_Robot"
VERSION : 0.1
   STRUCT
      status : "Fanuc_status";
      cmd : "Fanuc_cmd";
      grafcet : Struct
         int_Active_step : Int;
      END_STRUCT;
   END_STRUCT;
END_TYPE

TYPE "UR_Cobot"
VERSION : 0.1
   STRUCT
      status : "UR_1_T2O_State";
      cmd : Struct
         x_GoHome : Bool;
         x_Run_main_program : Bool;
         x_Hold : Bool;
         x_Reset_program : Bool;
         x_Reset_faults : Bool;
         x_Run_init_program : Bool;
      END_STRUCT;
      grafcet : Struct
         int_Active_step : Int;
      END_STRUCT;
      Registers : Struct
         Bit : "UR_5_T2O_BitRegisters";
         "Int" : "UR_6_T2O_IntRegisters";
         Float : "UR_7_T2O_FloatRegisters";
      END_STRUCT;
      Registers_Out_1 : "UR_9_O2T_Registers";
      Registers_Out_2 : "UR_9_O2T_Registers";
   END_STRUCT;
END_TYPE

TYPE "Fanuc_status"
VERSION : 0.1
   STRUCT
      x_Cmd_Enabled : Bool;
      x_Fault : Bool;
      x_Prog_Running : Bool;
      x_Snack : Bool;
      x_Teach_on : Bool;
      x_In_auto_mode : Bool;
      x_at_home_pos : Bool;
      x_libre_1 : Bool;
      x_Fin_prise : Bool;
      x_Fin_depose : Bool;
   END_STRUCT;
END_TYPE

TYPE "Fanuc_cmd"
VERSION : 0.1
   STRUCT
      x_IMSTP : Bool;
      x_Fault_reset : Bool;
      x_Start_Pns_strobe : Bool;
      x_Enable : Bool;
      x_PNS1 : Bool;
      x_PNS2 : Bool;
      x_Cicle_stop : Bool;
      x_Hold : Bool;
      x_Autor_Prise : Bool;
      x_Autor_Depose : Bool;
      x_GoHome : Bool;
      x_Avec_AGV : Bool;
   END_STRUCT;
END_TYPE

TYPE "Var_G120C_cmd"
VERSION : 0.1
   STRUCT
      Reserve01 : Bool;
      Reserve02 : Bool;
      PilotageParApi : Bool;
      InversionConsigne : Bool;
      Reserve03 : Bool;
      PotPlus : Bool;
      PotMoins : Bool;
      Reserve04 : Bool;
      Marche : Bool;
      Arret2 : Bool;
      Arret3 : Bool;
      DebloqFonctionnement : Bool;
      DebloqRampe : Bool;
      GelerGenerateurRampe : Bool;
      DebloqConsigne : Bool;
      AcquitDefaut : Bool;
      Consigne : Int;
   END_STRUCT;
END_TYPE

TYPE "Var_G120C_status"
VERSION : 0.1
   STRUCT
      EcartVitesse : Bool;
      CommandeDemander : Bool;
      VitesseMaxAtteinte : Bool;
      Limite : Bool;
      FreinMoteur : Bool;
      AlarmeSurchauffe : Bool;
      MoteurSensAvant : Bool;
      SurchargeMoteur : Bool;
      PretEnclenchement : Bool;
      PretFonctionnement : Bool;
      Fonctionnement_Debloq : Bool;
      DefautActif : Bool;
      Arret2Etat : Bool;
      Arret3Etat : Bool;
      BlocageActif : Bool;
      AlarmeActive : Bool;
      Vitesse : Int;
   END_STRUCT;
END_TYPE

TYPE "Var_G120C_data"
VERSION : 0.1
   STRUCT
      Status : "Var_G120C_status";
      Cmd : "Var_G120C_cmd";
   END_STRUCT;
END_TYPE

TYPE "GoFa_Status"
VERSION : 0.1
   STRUCT
      x_Collision_Avoidance : Bool;
      x_AU : Bool;
      x_Auto_On : Bool;
      x_Cycle_On : Bool;
      x_Rtc_Motors_On : Bool;
      x_Run_Chain_Ok : Bool;
      x_Home_Position : Bool;
      x_Colis_recuperé : Bool;
   END_STRUCT;
END_TYPE

TYPE "GoFa_cmd"
VERSION : 0.1
   STRUCT
      x_PP_vers_main : Bool;
      x_Motors_ON : Bool;
      x_Start : Bool;
      x_Motors_on_and_start : Bool;
      x_Stop : Bool;
      x_Stop_at_end_of_Instruction : Bool;
      x_Stop_at_end_of_cycle : Bool;
      x_Colis_pret : Bool;
   END_STRUCT;
END_TYPE

TYPE "Modbus_Read_Write"
VERSION : 0.1
   STRUCT
      Read : Array[0..31] of DInt;
      Write : Array[0..31] of DInt;
   END_STRUCT;
END_TYPE

// folder: UR_UDT

TYPE "UR__O2T_Robot"
VERSION : 0.1
   STRUCT
      "SSM: Speed slider fraction mask" : Bool;
      Reserved_1 : Bool;
      Reserved_2 : Bool;
      Reserved_3 : Bool;
      Reserved_4 : Bool;
      Reserved_5 : Bool;
      Reserved_6 : Bool;
      Reserved_7 : Bool;
      Reserved_8_15 : USInt;
      Reserved_16_31 : UInt;
      "Speed slider fraction" : Real;
   END_STRUCT;
END_TYPE

TYPE "UR__O2T_ints"
VERSION : 0.1
   STRUCT
      Register : Array[0..11] of DInt;
   END_STRUCT;
END_TYPE

TYPE "UR__O2T_floats"
VERSION : 0.1
   STRUCT
      Register : Array[0..11] of Real;
   END_STRUCT;
END_TYPE

TYPE "UR__O2T_IOs"
VERSION : 0.1
   STRUCT
      "Standard digital output mask" : USInt;
      "Configurable digital output mask" : USInt;
      "Standard digital outputs" : USInt;
      "Configurable digital outputs" : USInt;
      "AOM: Analog output mask" : USInt;
      "AOT: Analog output types" : USInt;
      "TDOM: Tool digital output mask" : USInt;
      "TDO: Tool digital output" : USInt;
      "Standard analog output" : Array[0..1] of Real;
   END_STRUCT;
END_TYPE

TYPE "UR__O2T_bits"
VERSION : 0.1
   STRUCT
      Register : Array[0..31] of Bool;
   END_STRUCT;
END_TYPE

TYPE "UR_9_O2T_Registers"
VERSION : 0.1
   STRUCT
      Bits : "UR__O2T_bits";
      Ints : "UR__O2T_ints";
      Floats : "UR__O2T_floats";
   END_STRUCT;
END_TYPE

TYPE "UR__T2O_IOs"
VERSION : 0.1
   STRUCT
      "Standard digital inputs" : USInt;
      "Configurable digital inputs" : USInt;
      "Standard digital outputs" : USInt;
      "Configurable digital outputs" : USInt;
      "Analog I/O types" : USInt;
      Reserved_8_15 : USInt;
      Reserved_16_31 : UInt;
      "Standard analog input [A or V]" : Array[0..1] of Real;
      "Standard analog output [A or V]" : Array[0..1] of Real;
      "I/O current [A]" : Real;
      "Euromap67 input bits" : Array[0..31] of Bool;
      "Euromap67 output bits" : Array[0..31] of Bool;
      "Euromap67 24V voltage" : Real;
      "Euromap67 24V current" : Real;
   END_STRUCT;
END_TYPE

TYPE "UR_8_O2T_Robot_IO"
VERSION : 0.1
   STRUCT
      Robot : "UR__O2T_Robot";
      IOs : "UR__O2T_IOs";
   END_STRUCT;
END_TYPE

TYPE "UR__T2O_Safety"
VERSION : 0.1
   STRUCT
      "Safety mode" : USInt;
      Reserved_1 : USInt;
      Reserved_2 : UInt;
      "NO: Is normal mode" : Bool;
      "RD: Is reduced mode" : Bool;
      "PS: Is protective stopped" : Bool;
      "RC: Is recovery mode" : Bool;
      "SS: Is safeguard stopped" : Bool;
      "SES: Is system emergency stopped" : Bool;
      "RES: Is robot emergency stopped" : Bool;
      "ES: Is emergency stopped" : Bool;
      "VL: Is violation" : Bool;
      "FT: Is fault" : Bool;
      "ST: Is stopped due to safety" : Bool;
      Reserved_11 : Bool;
      Reserved_12 : Bool;
      Reserved_13 : Bool;
      Reserved_14 : Bool;
      Reserved_15 : Bool;
      Reserved_16_31 : UInt;
   END_STRUCT;
END_TYPE

TYPE "UR__T2O_Robot"
VERSION : 0.1
   STRUCT
      "Controller major version" : USInt;
      "Controller minor version" : USInt;
      Reserved : UInt;
      "Robot mode" : USInt;
      "Real time machine seconds" : USInt;
      "Real time machine milliseconds" : UInt;
      "Real time machine minutes" : USInt;
      "Real time machine hours" : USInt;
      "Real time machine days" : UInt;
      "Robot current A" : Real;
      "PW: Is power on" : Bool;
      "PR: Is program running" : Bool;
      "TB: Is teach button pressed" : Bool;
      "PB: Is power button pressed" : Bool;
      Reserved_4 : Bool;
      Reserved_5 : Bool;
      Reserved_6 : Bool;
      Reserved_7 : Bool;
      Reserved_8_15 : USInt;
      Reserved_16_31 : UInt;
      "Speed slider fraction" : Real;
   END_STRUCT;
END_TYPE

TYPE "UR__T2O_Tool"
VERSION : 0.1
   STRUCT
      "Tool mode" : USInt;
      Reserved_7_15 : USInt;
      Reserved_16_31 : UInt;
      "TDI: Tool Digital Inputs" : USInt;
      "TDO: Tool Digital Outputs" : USInt;
      "TAIT: Tool Analog Input Types" : USInt;
      Reserved_24_31 : USInt;
      "Tool analog input [A or V]" : Array[0..1] of Real;
      "Tool output voltage [V]" : Real;
      "Tool current [A]" : Real;
   END_STRUCT;
END_TYPE

TYPE "UR_O2T"
VERSION : 0.1
   STRUCT
      "Robot IO" : "UR_8_O2T_Robot_IO";
      "Reg 1" : "UR_9_O2T_Registers";
      "Reg 2" : "UR_9_O2T_Registers";
   END_STRUCT;
END_TYPE

TYPE "UR_4_T2O_TCP"
VERSION : 0.1
   STRUCT
      "TCP Position (X,Y,Z) [m]" : Array[0..2] of Real;
      "TCP Position (RX,RY,RZ) [rad]" : Array[0..2] of Real;
      "TCP velocity (X,Y,Z) [m/s]" : Array[0..2] of Real;
      "TCP velocity (RX,RY,RZ) [rad/s]" : Array[0..2] of Real;
      "TCP force (X,Y,Z) [N]" : Array[0..2] of Real;
      "TCP torque (X,Y,Z) [Nm]" : Array[0..2] of Real;
      "TCP force scalar [N]" : Real;
   END_STRUCT;
END_TYPE

TYPE "UR_3_T2O_Joints"
VERSION : 0.1
   STRUCT
      "Joint position [rad]" : Array[0..5] of Real;
      "Joint velocity [rad/s]" : Array[0..5] of Real;
      "Joint current [A]" : Array[0..5] of Real;
      "Joint temperature [°C]" : Array[0..5] of Real;
      "Joint mode" : Array[0..5] of USInt;
      Reserved_9 : UInt;
   END_STRUCT;
END_TYPE

TYPE "UR_2_T2O_IO"
VERSION : 0.1
   STRUCT
      IOs : "UR__T2O_IOs";
      Tool : "UR__T2O_Tool";
   END_STRUCT;
END_TYPE

TYPE "UR_5_T2O_BitRegisters"
VERSION : 0.1
   STRUCT
      Register : Array[0..63] of Bool;
   END_STRUCT;
END_TYPE

TYPE "UR_1_T2O_State"
VERSION : 0.1
   STRUCT
      Robot : "UR__T2O_Robot";
      Safety : "UR__T2O_Safety";
   END_STRUCT;
END_TYPE

TYPE "UR_7_T2O_FloatRegisters"
VERSION : 0.1
   STRUCT
      Register : Array[0..23] of Real;
   END_STRUCT;
END_TYPE

TYPE "UR_6_T2O_IntRegisters"
VERSION : 0.1
   STRUCT
      Register : Array[0..23] of DInt;
   END_STRUCT;
END_TYPE

TYPE "UR_T2O"
VERSION : 0.1
   STRUCT
      State : "UR_1_T2O_State";
      IO : "UR_2_T2O_IO";
      Joints : "UR_3_T2O_Joints";
      TCP : "UR_4_T2O_TCP";
      Bits : "UR_5_T2O_BitRegisters";
      Ints : "UR_6_T2O_IntRegisters";
      Floats : "UR_7_T2O_FloatRegisters";
   END_STRUCT;
END_TYPE

// folder: 00_Donnees_globales

DATA_BLOCK "Voyants_HMI"   // DB4
{ S7_Optimized_Access := 'TRUE' }
VERSION : 0.1
   VAR
      x_VOY_Demo_pret : Bool;
      x_VOY_Tp_robot_pret : Bool;
      x_VOY_DCY : Bool;
      x_VOY_ACY : Bool;
      x_VOY_INIT : Bool;
      x_VOY_Init_requis_en_auto : Bool;
      x_VOY_AUTO_pret : Bool;
   END_VAR
BEGIN
END_DATA_BLOCK

DATA_BLOCK "Bits_Globaux"   // DB10
{ S7_Optimized_Access := 'TRUE' }
VERSION : 0.1
   VAR
      x_En_service : Bool;
      x_En_auto : Bool;
      x_En_manu : Bool;
      x_Defaut_bloquant : Bool;
      x_Defaut_non_bloquant : Bool;
      x_Demo_Hippo_en_cours : Bool;
      x_Init_glob_OK : Bool;
      x_Init_en_cours : Bool;
      x_Dmd_Init_robot : Bool;
      x_Tp_Robots_en_cours : Bool;
      x_Robots_en_AUTO : Bool;
      x_En_cycle_auto : Bool;
   END_VAR
BEGIN
END_DATA_BLOCK

DATA_BLOCK "Tch_HMI"   // DB11
{ S7_Optimized_Access := 'TRUE' }
VERSION : 0.1
   VAR
      Tch_Dcy : Bool;
      Tch_Acy : Bool;
      Tch_Acquit : Bool;
      Tch_Init : Bool;
      Tch_Tp_Robot : Bool;
      Tch_Demo : Bool;
      Tch_Manu : Array[0..100] of Bool;
   END_VAR
BEGIN
   // Tch_Manu[62] : Marche convoyeur CV01
   // Tch_Manu[63] : Arret convoyeur CV01
   // Tch_Manu[64] : Marche convoyeur CV02
   // Tch_Manu[65] : Arret convoyeur CV02
   // Tch_Manu[66] : Marche convoyeur CV03
   // Tch_Manu[67] : Arret convoyeur CV03
   // Tch_Manu[92] : Envoi trigger vision Keyence
END_DATA_BLOCK

DATA_BLOCK "Défauts"   // DB13
{ S7_Optimized_Access := 'FALSE' }
VERSION : 0.1
   VAR
      Defauts : Array[0..100] of Bool;
      Def_Canal01 : Int;
      Def_Canal02 : Int;
      Def_Canal03 : Int;
   END_VAR
BEGIN
END_DATA_BLOCK

DATA_BLOCK "Parametres"   // DB18
{ S7_Optimized_Access := 'TRUE' }
VERSION : 0.1
   VAR RETAIN
      Convoyeurs : Struct
         Auto : Struct
            i_Vitesse_C01 : Int := 400;
            i_Vitesse_C02 : Int := 400;
            i_Vitesse_C03 : Int := 400;
         END_STRUCT;
         Manu : Struct
            i_Vitesse_manu_C01 : Int := 400;
            i_Vitesse_manu_C02 : Int := 400;
            i_Vitesse_manu_C03 : Int := 400;
         END_STRUCT;
      END_STRUCT;
   END_VAR
BEGIN
END_DATA_BLOCK

DATA_BLOCK "Defauts_DB"   // DB32
{ S7_Optimized_Access := 'TRUE' }
VERSION : 0.1
// stored: InstanceOfName Defauts
"Defauts"
BEGIN
   "Erreur elevateur hippodrome"[0] := 'Defaut elevateur hippodrome';
   "Erreur elevateur hippodrome"[1] := 'L elevateur n a pas atteint la position requise';
END_DATA_BLOCK

// folder: 1_Imprimantes_3D

DATA_BLOCK "DB_Imprimantes"   // DB2
{ S7_Optimized_Access := 'TRUE' }
VERSION : 0.1
   VAR
      Imprimante : Array[1..4] of "Imprimante3D";
   END_VAR
BEGIN
   Imprimante[1].Printer_ID := 1;
   Imprimante[2].Printer_ID := 2;
   Imprimante[3].Printer_ID := 3;
   Imprimante[4].Printer_ID := 4;
   // Imprimante[1] : Données imprimante n°1
   // Imprimante[2] : Données imprimante n°2
   // Imprimante[3] : Données imprimante n°3
   // Imprimante[4] : Données imprimante n°4
END_DATA_BLOCK

// folder: 2-Hippodrome/Convoyeurs

DATA_BLOCK "DB_Convoyeurs_Hipp"   // DB1
{ S7_Optimized_Access := 'TRUE' }
VERSION : 0.1
   VAR
      Convoyeur : Array[1..4] of "Convoyeur_Hipp";
   END_VAR
BEGIN
END_DATA_BLOCK

DATA_BLOCK "21_Gestion_Convoyeurs_hippodrome_DB"   // DB15
{ S7_Optimized_Access := 'TRUE' }
VERSION : 0.1
// stored: InstanceOfName 21_Gestion_Convoyeurs_hippodrome
"21_Gestion_Convoyeurs_hippodrome"
BEGIN
END_DATA_BLOCK

// folder: 2-Hippodrome/Stations de travail

DATA_BLOCK "DB_Stations"   // DB3
{ S7_Optimized_Access := 'TRUE' }
VERSION : 0.1
   VAR
      Station : Array[1..7] of "Station_Hipp";
   END_VAR
BEGIN
   Station[1].Num_station := 1;
   Station[2].Num_station := 2;
   Station[3].Num_station := 3;
   Station[4].Num_station := 4;
   Station[5].Num_station := 5;
   Station[6].Num_station := 6;
   Station[7].Num_station := 7;
END_DATA_BLOCK

DATA_BLOCK "22-Gestion_stations_DB"   // DB16
{ S7_Optimized_Access := 'TRUE' }
VERSION : 0.1
// stored: InstanceOfName 22-Gestion_stations
"22-Gestion_stations"
BEGIN
END_DATA_BLOCK

// folder: 3_Controle vision

DATA_BLOCK "DB_Projet_Vision"   // DB14
{ S7_Optimized_Access := 'TRUE' }
VERSION : 0.1
   VAR
      Validation : Bool;
      Entree_FIFO : Int;
      Sortie_FIFO : Int;
      "M" : Bool;
   END_VAR
BEGIN
END_DATA_BLOCK

DATA_BLOCK "DB_FIFO"   // DB19
{ S7_Optimized_Access := 'TRUE' }
VERSION : 0.1
// stored: InstanceOfName FIFO
"FIFO"
BEGIN
END_DATA_BLOCK

DATA_BLOCK "31_Keyence_Camera_DB"   // DB23
{ S7_Optimized_Access := 'TRUE' }
VERSION : 0.1
// stored: InstanceOfName 31_Keyence_Camera
"31_Keyence_Camera"
BEGIN
END_DATA_BLOCK

DATA_BLOCK "32_Cmd_porte_vision_DB"   // DB24
{ S7_Optimized_Access := 'TRUE' }
VERSION : 0.1
// stored: InstanceOfName 32_Cmd_porte_vision
"32_Cmd_porte_vision"
BEGIN
END_DATA_BLOCK

DATA_BLOCK "Vision_Keyence"   // DB73
{ S7_Optimized_Access := 'TRUE' }
VERSION : 0.1
   VAR
      Step_cycle : Int;
      Trans : Struct
         "00" : Bool;
         "01" : Bool;
         "12" : Bool;
         "23" : Bool;
         "34" : Bool;
         "45" : Bool;
         "56" : Bool;
         "67" : Bool;
         "78" : Bool;
         "89" : Bool;
      END_STRUCT;
   END_VAR
BEGIN
END_DATA_BLOCK

// folder: 4_UR10_R4

DATA_BLOCK "40_UR_R4_DB"   // DB12
{ S7_Optimized_Access := 'TRUE' }
VERSION : 0.1
// stored: InstanceOfName 40_UR_R4
"40_UR_R4"
BEGIN
END_DATA_BLOCK

// folder: 5-Cellule_conditionnement/Convoyeurs

DATA_BLOCK "Gestion_Convoyeurs_DB"   // DB6
{ S7_Optimized_Access := 'TRUE' }
VERSION : 0.1
// stored: InstanceOfName Gestion_Convoyeurs
"Gestion_Convoyeurs"
BEGIN
END_DATA_BLOCK

DATA_BLOCK "DB_Variateurs"   // DB17
{ S7_Optimized_Access := 'FALSE' }
VERSION : 0.1
   VAR
      ConvoyeurC01 : "Var_G120C_data";
      ConvoyeurC02 : "Var_G120C_data";
      ConvoyeurC03 : "Var_G120C_data";
   END_VAR
BEGIN
END_DATA_BLOCK

// folder: 5-Cellule_conditionnement/Fanuc_R1

DATA_BLOCK "Fanuc_R1_DB"   // DB7
{ S7_Optimized_Access := 'TRUE' }
VERSION : 0.1
// stored: InstanceOfName Fanuc_R1
"Fanuc_R1"
BEGIN
END_DATA_BLOCK

// folder: 5-Cellule_conditionnement/Fanuc_R2

DATA_BLOCK "Fanuc_R2_DB"   // DB8
{ S7_Optimized_Access := 'TRUE' }
VERSION : 0.1
// stored: InstanceOfName Fanuc_R2
"Fanuc_R2"
BEGIN
END_DATA_BLOCK

// folder: 5-Cellule_conditionnement/GoFa_ABB_R3

DATA_BLOCK "GoFa_R3_FB_DB"   // DB25
{ S7_Optimized_Access := 'TRUE' }
VERSION : 0.1
// stored: InstanceOfName GoFa_R3_FB
"GoFa_R3_FB"
BEGIN
END_DATA_BLOCK

// folder: 6_UR10_R5

DATA_BLOCK "60_UR_R5_DB"   // DB9
{ S7_Optimized_Access := 'TRUE' }
VERSION : 0.1
// stored: InstanceOfName 60_UR_R5
"60_UR_R5"
BEGIN
END_DATA_BLOCK

// folder: 7_AGVs

DATA_BLOCK "AGVs_Modbus_Write_COM_DB"   // DB26
{ S7_Optimized_Access := 'TRUE' }
VERSION : 0.1
// stored: InstanceOfName AGVs_Modbus_Write_COM
"AGVs_Modbus_Write_COM"
BEGIN
END_DATA_BLOCK

DATA_BLOCK "AGVs_Modbus_Read_COM_DB"   // DB27
{ S7_Optimized_Access := 'TRUE' }
VERSION : 0.1
// stored: InstanceOfName AGVs_Modbus_Read_COM
"AGVs_Modbus_Read_COM"
BEGIN
END_DATA_BLOCK

DATA_BLOCK "HR_Modbus_AGV"   // DB28
{ S7_Optimized_Access := 'FALSE' }
VERSION : 0.1
   VAR
      AGV1 : "Modbus_Read_Write";
      AGV2 : "Modbus_Read_Write";
   END_VAR
BEGIN
   AGV1.Write[0] := 0;   // Etat_boucle_recup_GC_ABB
   // AGV1.Read[0] : Etat_boucle_recup_GC_ABB
   // AGV1.Read[1] : Etat_boucle_recup_PC_UR4
   // AGV1.Read[2] : Etat_boucle_recup_GC_UR5
   // AGV1.Read[3] : GO_HOME_1
   // AGV1.Read[4] : GO_HOME_2
   // AGV1.Read[5] : Charge_needed
   // AGV1.Write[1] : Etat_boucle_recup_PC_UR4
   // AGV1.Write[2] : Etat_boucle_recup_GC_UR5
   // AGV1.Write[3] : GO_HOME_1
   // AGV1.Write[4] : GO_HOME_2
   // AGV1.Write[5] : Charge_needed
END_DATA_BLOCK

DATA_BLOCK "AGV_1_DB"   // DB29
{ S7_Optimized_Access := 'TRUE' }
VERSION : 0.1
// stored: InstanceOfName AGV_1
"AGV_1"
BEGIN
END_DATA_BLOCK

DATA_BLOCK "Connection_params"   // DB30
{ S7_Optimized_Access := 'TRUE' }
VERSION : 0.1
   VAR RETAIN
      AGV_1_read : TCON_IP_v4;
   END_VAR
   VAR
      AGV_1_write : TCON_IP_v4;
   END_VAR
   VAR RETAIN
      AGV_2_read : TCON_IP_v4;
   END_VAR
   VAR
      AGV_2_write : TCON_IP_v4;
   END_VAR
BEGIN
   AGV_1_read.RemoteAddress.ADDR[1] := 172;
   AGV_1_read.RemoteAddress.ADDR[2] := 16;
   AGV_1_read.RemoteAddress.ADDR[3] := 1;
   AGV_1_read.RemoteAddress.ADDR[4] := 190;
   AGV_1_read.RemotePort := 502;
   AGV_1_read.LocalPort := 0;
   AGV_1_read.ID := 1;
   AGV_1_read.ConnectionType := 11;
   AGV_1_read.ActiveEstablished := 1;
   AGV_1_read.InterfaceId := 64;
   AGV_2_read.InterfaceId := 64;
   AGV_2_read.ID := 3;
   AGV_2_read.ConnectionType := 11;
   AGV_2_read.ActiveEstablished := 1;
   AGV_2_read.RemoteAddress.ADDR[1] := 172;
   AGV_2_read.RemoteAddress.ADDR[2] := 16;
   AGV_2_read.RemoteAddress.ADDR[3] := 1;
   AGV_2_read.RemoteAddress.ADDR[4] := 191;
   AGV_2_read.RemotePort := 502;
   AGV_2_read.LocalPort := 0;
   AGV_1_write.InterfaceId := 64;
   AGV_1_write.ID := 2;
   AGV_1_write.ConnectionType := 11;
   AGV_1_write.ActiveEstablished := 1;
   AGV_1_write.RemotePort := 502;
   AGV_1_write.LocalPort := 0;
   AGV_1_write.RemoteAddress.ADDR[1] := 172;
   AGV_1_write.RemoteAddress.ADDR[2] := 16;
   AGV_1_write.RemoteAddress.ADDR[3] := 1;
   AGV_1_write.RemoteAddress.ADDR[4] := 190;
   AGV_2_write.InterfaceId := 64;
   AGV_2_write.ID := 4;
   AGV_2_write.ConnectionType := 11;
   AGV_2_write.ActiveEstablished := 1;
   AGV_2_write.LocalPort := 0;
   AGV_2_write.RemoteAddress.ADDR[1] := 172;
   AGV_2_write.RemoteAddress.ADDR[2] := 16;
   AGV_2_write.RemoteAddress.ADDR[3] := 1;
   AGV_2_write.RemoteAddress.ADDR[4] := 191;
   AGV_2_write.RemotePort := 502;
END_DATA_BLOCK

DATA_BLOCK "AGV_2_DB"   // DB31
{ S7_Optimized_Access := 'TRUE' }
VERSION : 0.1
// stored: InstanceOfName AGV_2
"AGV_2"
BEGIN
END_DATA_BLOCK

// folder: System blocks/Program resources

DATA_BLOCK "Init_Timer"   // DB5
{ S7_Optimized_Access := 'TRUE' }
AUTHOR : Simatic
FAMILY : IEC
NAME : IEC_TMR
VERSION : 1.0
// stored: InstanceOfName IEC_TIMER
"IEC_TIMER"
BEGIN
END_DATA_BLOCK

DATA_BLOCK "IEC_Counter_0_DB"   // DB20
{ S7_Optimized_Access := 'TRUE' }
AUTHOR : Simatic
FAMILY : IEC
NAME : CNTR
VERSION : 1.0
// stored: InstanceOfName IEC_COUNTER
"IEC_COUNTER"
BEGIN
END_DATA_BLOCK

DATA_BLOCK "Timer_Test_Fanuc"   // DB21
{ S7_Optimized_Access := 'TRUE' }
AUTHOR : Simatic
FAMILY : IEC
NAME : IEC_TMR
VERSION : 1.0
// stored: InstanceOfName IEC_TIMER
"IEC_TIMER"
BEGIN
END_DATA_BLOCK

DATA_BLOCK "Test_Sncak"   // DB22
{ S7_Optimized_Access := 'TRUE' }
AUTHOR : Simatic
FAMILY : IEC
NAME : IEC_TMR
VERSION : 1.0
// stored: InstanceOfName IEC_TIMER
"IEC_TIMER"
BEGIN
END_DATA_BLOCK

// folder: (top level)

ORGANIZATION_BLOCK "Main"   // OB1, LAD, ProgramCycle
TITLE = "Main Program Sweep (Cycle)"
{ S7_Optimized_Access := 'TRUE' }
VERSION : 0.1
   VAR_INPUT
      Initial_Call : Bool;   // Initial call of this OB
      Remanence : Bool;   // =True, if remanent data are available
   END_VAR
   VAR_TEMP   // added for the SCL form of the ladder/FBD networks
      _w1 : Bool;
   END_VAR
BEGIN

REGION Network 1: Copie IOs Equipements
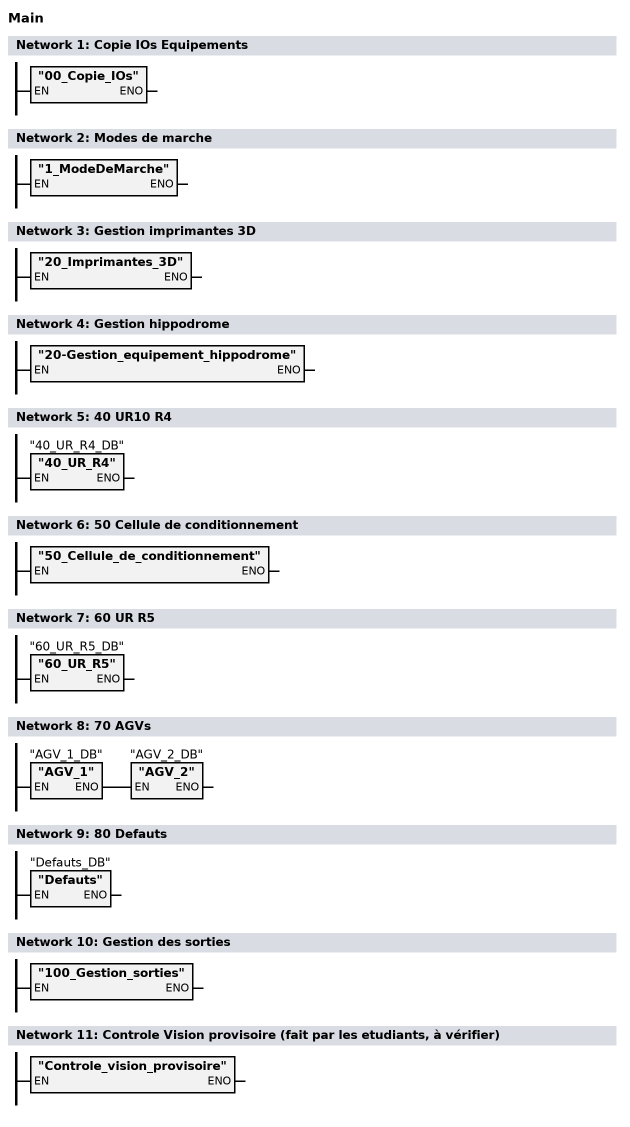
   RUNG wire#powerrail
      "00_Copie_IOs"()
   END_RUNG
   // the same network as SCL:
   "00_Copie_IOs"();
END_REGION

REGION Network 2: Modes de marche
   RUNG wire#powerrail
      "1_ModeDeMarche"()
   END_RUNG
   // the same network as SCL:
   "1_ModeDeMarche"();
END_REGION

REGION Network 3: Gestion imprimantes 3D
   RUNG wire#powerrail
      "20_Imprimantes_3D"()
   END_RUNG
   // the same network as SCL:
   "20_Imprimantes_3D"();
END_REGION

REGION Network 4: Gestion hippodrome
   RUNG wire#powerrail
      "20-Gestion_equipement_hippodrome"()
   END_RUNG
   // the same network as SCL:
   "20-Gestion_equipement_hippodrome"();
END_REGION

REGION Network 5: 40 UR10 R4
   RUNG wire#powerrail
      "40_UR_R4_DB"()
   END_RUNG
   // the same network as SCL:
   "40_UR_R4_DB"();   // "40_UR_R4"
END_REGION

REGION Network 6: 50 Cellule de conditionnement
   RUNG wire#powerrail
      "50_Cellule_de_conditionnement"()
   END_RUNG
   // the same network as SCL:
   "50_Cellule_de_conditionnement"();
END_REGION

REGION Network 7: 60 UR R5
   RUNG wire#powerrail
      "60_UR_R5_DB"()
   END_RUNG
   // the same network as SCL:
   "60_UR_R5_DB"();   // "60_UR_R5"
END_REGION

REGION Network 8: 70 AGVs
   RUNG wire#powerrail
      "AGV_1_DB"()
      "AGV_2_DB"()
   END_RUNG
   // the same network as SCL:
   "AGV_1_DB"(ENO => #_w1);   // "AGV_1"
   IF #_w1 THEN
       "AGV_2_DB"();   // "AGV_2"
   END_IF;
END_REGION

REGION Network 9: 80 Defauts
   RUNG wire#powerrail
      "Defauts_DB"()
   END_RUNG
   // the same network as SCL:
   "Defauts_DB"();   // "Defauts"
END_REGION

REGION Network 10: Gestion des sorties
   RUNG wire#powerrail
      "100_Gestion_sorties"()
   END_RUNG
   // the same network as SCL:
   "100_Gestion_sorties"();
END_REGION

REGION Network 11: Controle Vision provisoire (fait par les etudiants, à vérifier)
   RUNG wire#powerrail
      "Controle_vision_provisoire"()
   END_RUNG
   // the same network as SCL:
   "Controle_vision_provisoire"();
END_REGION
END_ORGANIZATION_BLOCK

// folder: 00_Donnees_globales

FUNCTION "1_ModeDeMarche" : Void   // FC1, LAD
{ S7_Optimized_Access := 'TRUE' }
VERSION : 0.1
BEGIN

REGION Network 1: Mise en Service
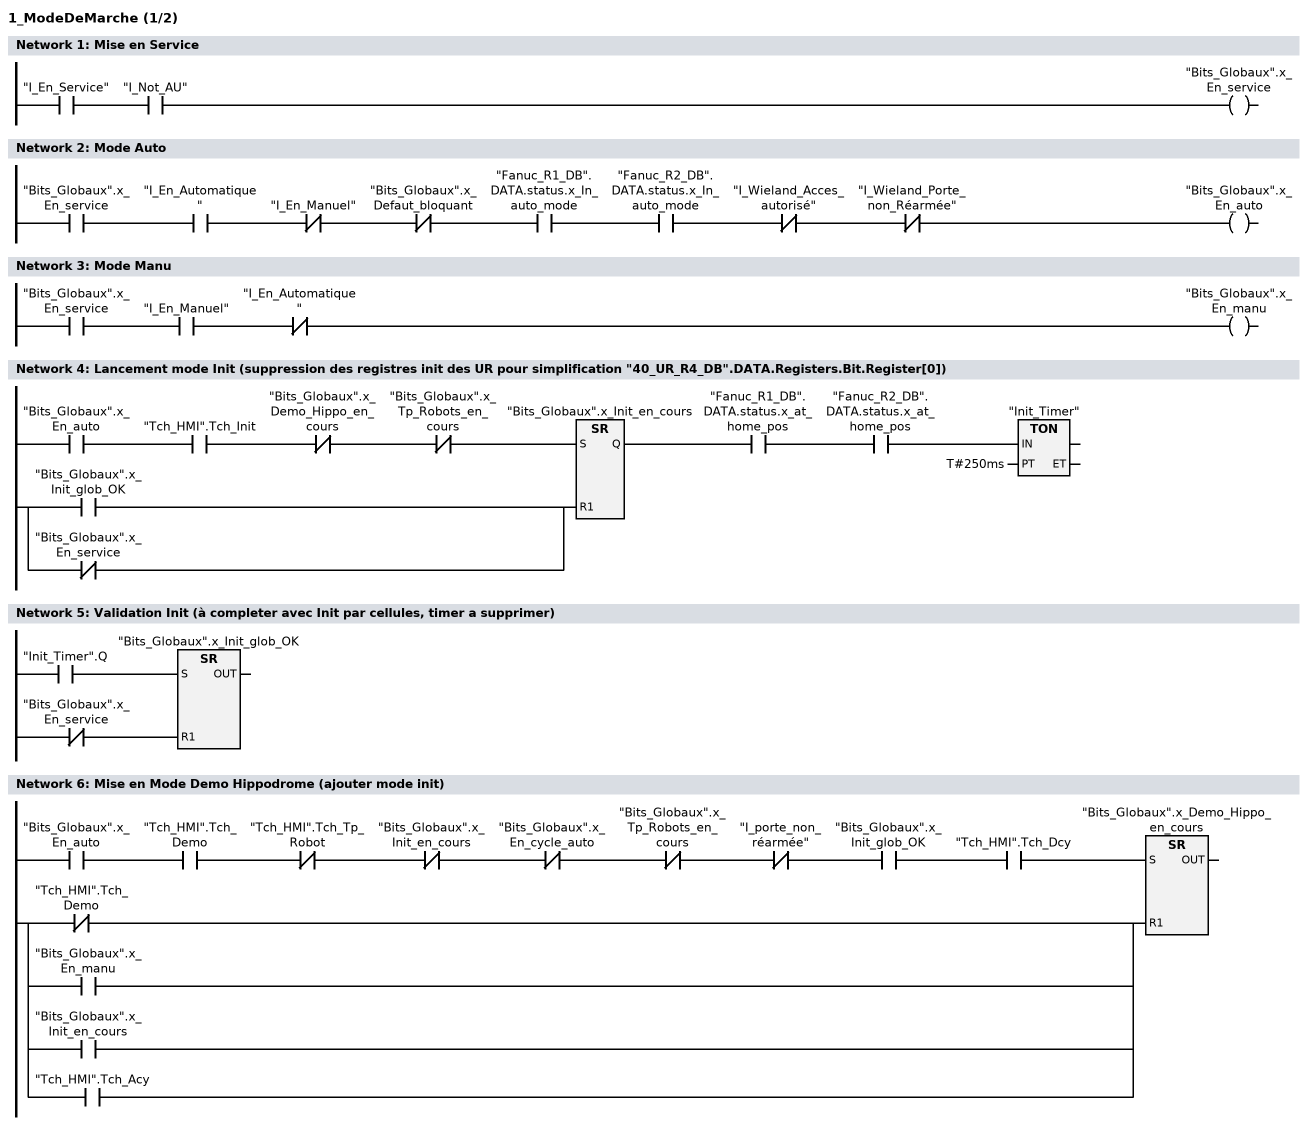
   RUNG wire#powerrail
      Contact( "I_En_Service" )
      Contact( "I_Not_AU" )
      Coil( "Bits_Globaux".x_En_service )
   END_RUNG
   // the same network as SCL:
   "Bits_Globaux".x_En_service := "I_En_Service" AND "I_Not_AU";
END_REGION

REGION Network 2: Mode Auto
   RUNG wire#powerrail
      Contact( "Bits_Globaux".x_En_service )
      Contact( "I_En_Automatique" )
      I_Contact( "I_En_Manuel" )
      I_Contact( "Bits_Globaux".x_Defaut_bloquant )
      Contact( "Fanuc_R1_DB".DATA.status.x_In_auto_mode )
      Contact( "Fanuc_R2_DB".DATA.status.x_In_auto_mode )
      I_Contact( "I_Wieland_Acces_autorisé" )
      I_Contact( "I_Wieland_Porte_non_Réarmée" )
      Coil( "Bits_Globaux".x_En_auto )
   END_RUNG
   // the same network as SCL:
   "Bits_Globaux".x_En_auto := "Bits_Globaux".x_En_service AND "I_En_Automatique" AND NOT "I_En_Manuel" AND NOT "Bits_Globaux".x_Defaut_bloquant AND "Fanuc_R1_DB".DATA.status.x_In_auto_mode AND "Fanuc_R2_DB".DATA.status.x_In_auto_mode AND NOT "I_Wieland_Acces_autorisé" AND NOT "I_Wieland_Porte_non_Réarmée";
END_REGION

REGION Network 3: Mode Manu
   RUNG wire#powerrail
      Contact( "Bits_Globaux".x_En_service )
      Contact( "I_En_Manuel" )
      I_Contact( "I_En_Automatique" )
      Coil( "Bits_Globaux".x_En_manu )
   END_RUNG
   // the same network as SCL:
   "Bits_Globaux".x_En_manu := "Bits_Globaux".x_En_service AND "I_En_Manuel" AND NOT "I_En_Automatique";
END_REGION

REGION Network 4: Lancement mode Init (suppression des registres init des UR pour simplification "40_UR_R4_DB".DATA.Registers.Bit.Register[0])
   IF "Bits_Globaux".x_En_auto AND "Tch_HMI".Tch_Init AND NOT "Bits_Globaux".x_Demo_Hippo_en_cours AND NOT "Bits_Globaux".x_Tp_Robots_en_cours THEN
       "Bits_Globaux".x_Init_en_cours := TRUE;   // SR flip-flop
   END_IF;
   IF "Bits_Globaux".x_Init_glob_OK OR NOT "Bits_Globaux".x_En_service THEN
       "Bits_Globaux".x_Init_en_cours := FALSE;
   END_IF;
   "Init_Timer".TON(IN := "Bits_Globaux".x_Init_en_cours AND "Fanuc_R1_DB".DATA.status.x_at_home_pos AND "Fanuc_R2_DB".DATA.status.x_at_home_pos,
                    PT := T#250ms);
END_REGION

REGION Network 5: Validation Init (à completer avec Init par cellules, timer a supprimer)
   RUNG wire#powerrail
      Contact( "Init_Timer".Q )
      S_SR(operand := "Bits_Globaux".x_Init_glob_OK, r1 := wire#w1)
   END_RUNG
   RUNG wire#powerrail
      I_Contact( "Bits_Globaux".x_En_service )
   END_RUNG wire#w1
   // the same network as SCL:
   IF "Init_Timer".Q THEN
       "Bits_Globaux".x_Init_glob_OK := TRUE;   // SR flip-flop
   END_IF;
   IF NOT "Bits_Globaux".x_En_service THEN "Bits_Globaux".x_Init_glob_OK := FALSE; END_IF;
END_REGION

REGION Network 6: Mise en Mode Demo Hippodrome (ajouter mode init)
   RUNG wire#powerrail
      Contact( "Bits_Globaux".x_En_auto )
      Contact( "Tch_HMI".Tch_Demo )
      I_Contact( "Tch_HMI".Tch_Tp_Robot )
      I_Contact( "Bits_Globaux".x_Init_en_cours )
      I_Contact( "Bits_Globaux".x_En_cycle_auto )
      I_Contact( "Bits_Globaux".x_Tp_Robots_en_cours )
      I_Contact( "I_porte_non_réarmée" )
      Contact( "Bits_Globaux".x_Init_glob_OK )
      Contact( "Tch_HMI".Tch_Dcy )
      S_SR(operand := "Bits_Globaux".x_Demo_Hippo_en_cours, r1 := wire#w1)
   END_RUNG
   RUNG wire#powerrail
      I_Contact( "Tch_HMI".Tch_Demo )
   END_RUNG wire#w1
   RUNG wire#powerrail
      Contact( "Bits_Globaux".x_En_manu )
   END_RUNG wire#w1
   RUNG wire#powerrail
      Contact( "Bits_Globaux".x_Init_en_cours )
   END_RUNG wire#w1
   RUNG wire#powerrail
      Contact( "Tch_HMI".Tch_Acy )
   END_RUNG wire#w1
   // the same network as SCL:
   IF "Bits_Globaux".x_En_auto AND "Tch_HMI".Tch_Demo AND NOT "Tch_HMI".Tch_Tp_Robot AND NOT "Bits_Globaux".x_Init_en_cours AND NOT "Bits_Globaux".x_En_cycle_auto AND NOT "Bits_Globaux".x_Tp_Robots_en_cours AND NOT "I_porte_non_réarmée" AND "Bits_Globaux".x_Init_glob_OK AND "Tch_HMI".Tch_Dcy THEN
       "Bits_Globaux".x_Demo_Hippo_en_cours := TRUE;   // SR flip-flop
   END_IF;
   IF NOT "Tch_HMI".Tch_Demo OR "Bits_Globaux".x_En_manu OR "Bits_Globaux".x_Init_en_cours OR "Tch_HMI".Tch_Acy THEN
       "Bits_Globaux".x_Demo_Hippo_en_cours := FALSE;
   END_IF;
END_REGION

REGION Network 7: Mise en Mode TP Robot
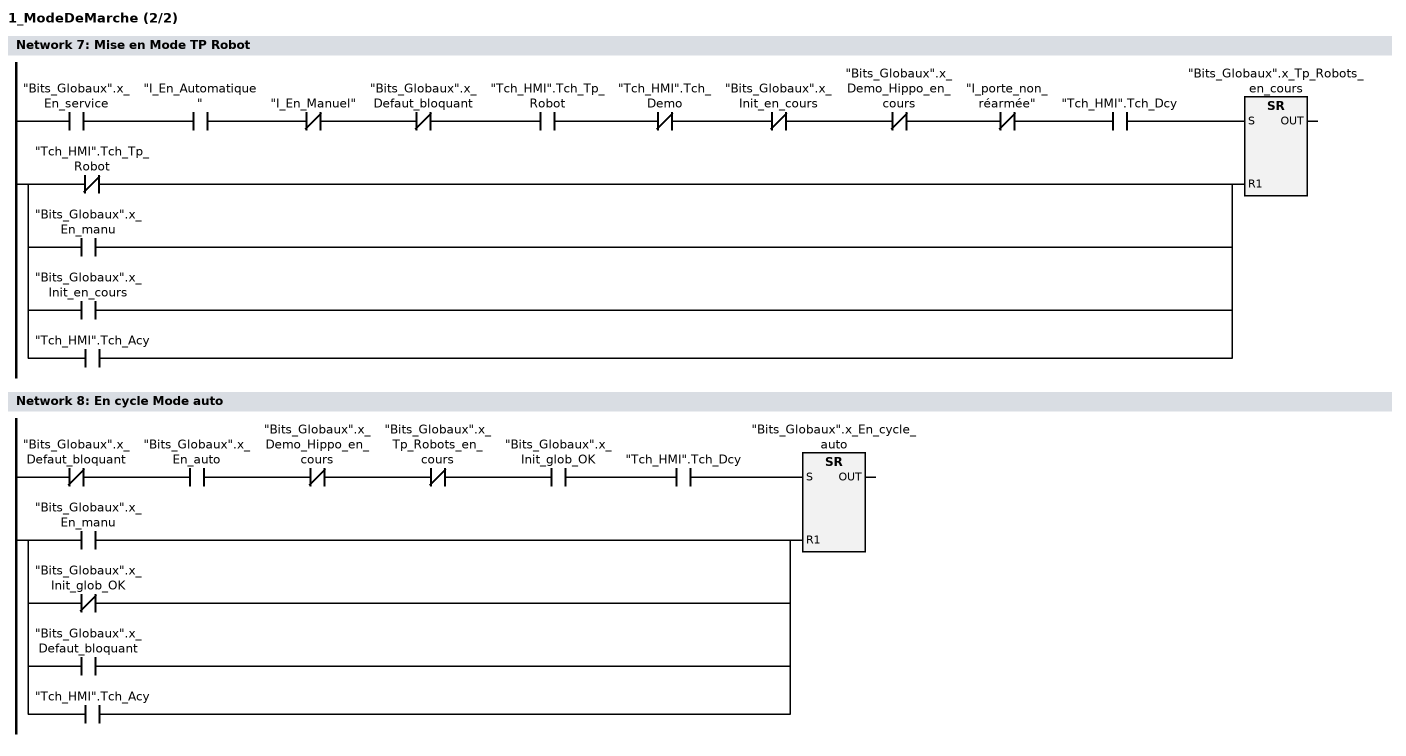
   RUNG wire#powerrail
      Contact( "Bits_Globaux".x_En_service )
      Contact( "I_En_Automatique" )
      I_Contact( "I_En_Manuel" )
      I_Contact( "Bits_Globaux".x_Defaut_bloquant )
      Contact( "Tch_HMI".Tch_Tp_Robot )
      I_Contact( "Tch_HMI".Tch_Demo )
      I_Contact( "Bits_Globaux".x_Init_en_cours )
      I_Contact( "Bits_Globaux".x_Demo_Hippo_en_cours )
      I_Contact( "I_porte_non_réarmée" )
      Contact( "Tch_HMI".Tch_Dcy )
      S_SR(operand := "Bits_Globaux".x_Tp_Robots_en_cours, r1 := wire#w1)
   END_RUNG
   RUNG wire#powerrail
      I_Contact( "Tch_HMI".Tch_Tp_Robot )
   END_RUNG wire#w1
   RUNG wire#powerrail
      Contact( "Bits_Globaux".x_En_manu )
   END_RUNG wire#w1
   RUNG wire#powerrail
      Contact( "Bits_Globaux".x_Init_en_cours )
   END_RUNG wire#w1
   RUNG wire#powerrail
      Contact( "Tch_HMI".Tch_Acy )
   END_RUNG wire#w1
   // the same network as SCL:
   IF "Bits_Globaux".x_En_service AND "I_En_Automatique" AND NOT "I_En_Manuel" AND NOT "Bits_Globaux".x_Defaut_bloquant AND "Tch_HMI".Tch_Tp_Robot AND NOT "Tch_HMI".Tch_Demo AND NOT "Bits_Globaux".x_Init_en_cours AND NOT "Bits_Globaux".x_Demo_Hippo_en_cours AND NOT "I_porte_non_réarmée" AND "Tch_HMI".Tch_Dcy THEN
       "Bits_Globaux".x_Tp_Robots_en_cours := TRUE;   // SR flip-flop
   END_IF;
   IF NOT "Tch_HMI".Tch_Tp_Robot OR "Bits_Globaux".x_En_manu OR "Bits_Globaux".x_Init_en_cours OR "Tch_HMI".Tch_Acy THEN
       "Bits_Globaux".x_Tp_Robots_en_cours := FALSE;
   END_IF;
END_REGION

REGION Network 8: En cycle Mode auto
   RUNG wire#powerrail
      I_Contact( "Bits_Globaux".x_Defaut_bloquant )
      Contact( "Bits_Globaux".x_En_auto )
      I_Contact( "Bits_Globaux".x_Demo_Hippo_en_cours )
      I_Contact( "Bits_Globaux".x_Tp_Robots_en_cours )
      Contact( "Bits_Globaux".x_Init_glob_OK )
      Contact( "Tch_HMI".Tch_Dcy )
      S_SR(operand := "Bits_Globaux".x_En_cycle_auto, r1 := wire#w1)
   END_RUNG
   RUNG wire#powerrail
      Contact( "Bits_Globaux".x_En_manu )
   END_RUNG wire#w1
   RUNG wire#powerrail
      I_Contact( "Bits_Globaux".x_Init_glob_OK )
   END_RUNG wire#w1
   RUNG wire#powerrail
      Contact( "Bits_Globaux".x_Defaut_bloquant )
   END_RUNG wire#w1
   RUNG wire#powerrail
      Contact( "Tch_HMI".Tch_Acy )
   END_RUNG wire#w1
   // the same network as SCL:
   IF NOT "Bits_Globaux".x_Defaut_bloquant AND "Bits_Globaux".x_En_auto AND NOT "Bits_Globaux".x_Demo_Hippo_en_cours AND NOT "Bits_Globaux".x_Tp_Robots_en_cours AND "Bits_Globaux".x_Init_glob_OK AND "Tch_HMI".Tch_Dcy THEN
       "Bits_Globaux".x_En_cycle_auto := TRUE;   // SR flip-flop
   END_IF;
   IF "Bits_Globaux".x_En_manu OR NOT "Bits_Globaux".x_Init_glob_OK OR "Bits_Globaux".x_Defaut_bloquant OR "Tch_HMI".Tch_Acy THEN
       "Bits_Globaux".x_En_cycle_auto := FALSE;
   END_IF;
END_REGION
END_FUNCTION

FUNCTION "00_Copie_IOs" : Void   // FC6, LAD
{ S7_Optimized_Access := 'TRUE' }
VERSION : 0.1
BEGIN

REGION Network 1: Copie ETAT UR R4
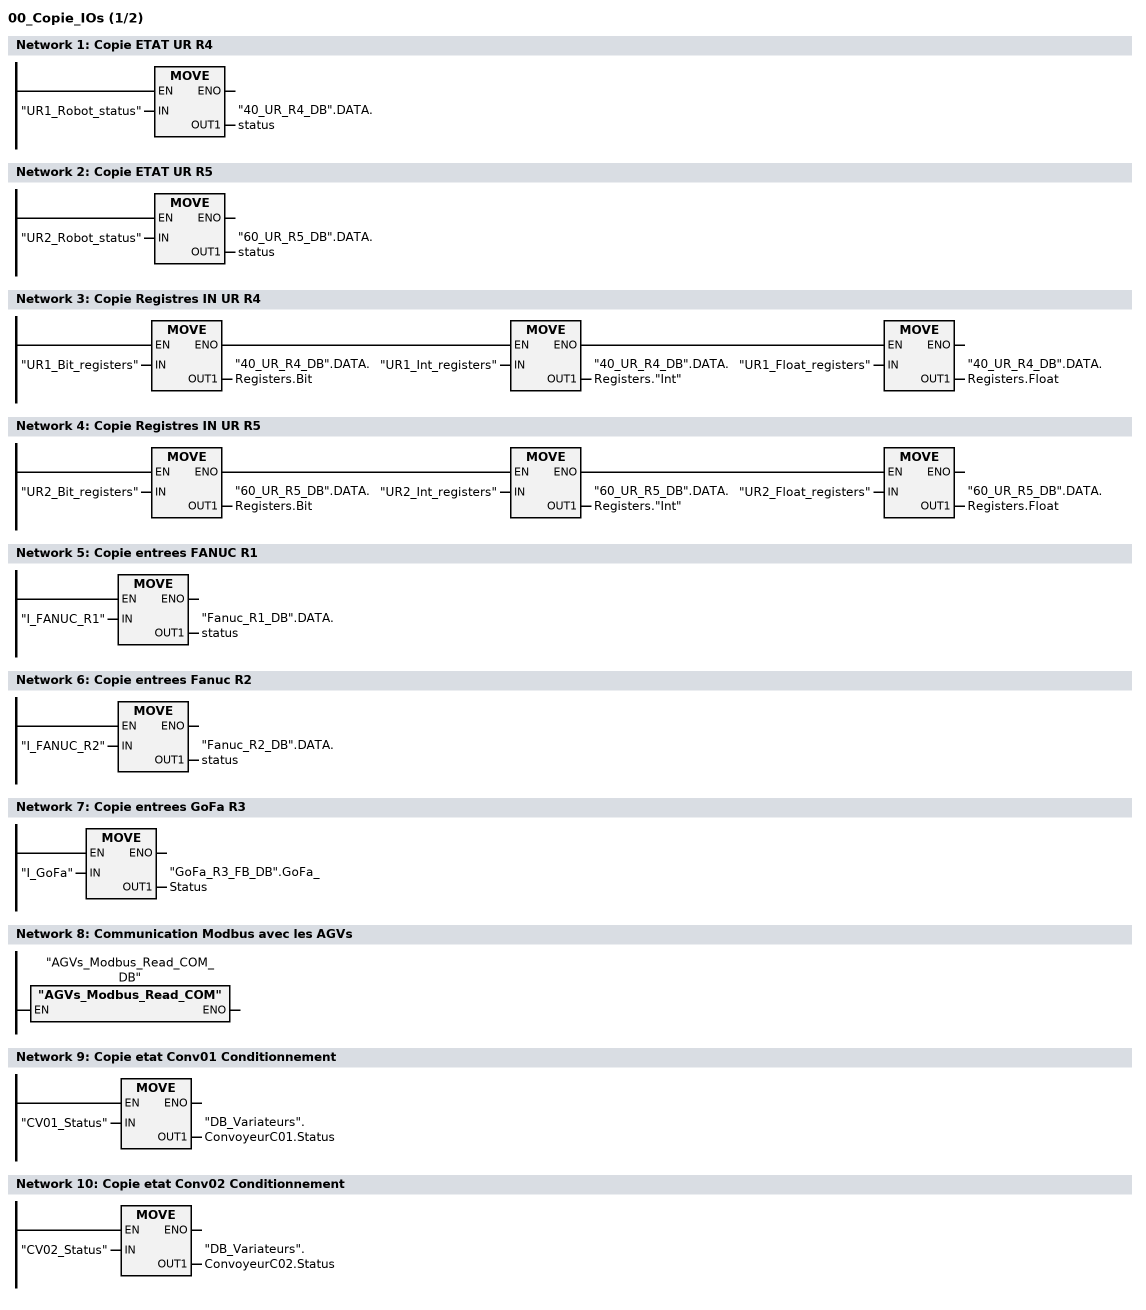
   RUNG wire#powerrail
      Move(in := "UR1_Robot_status", out1 => "40_UR_R4_DB".DATA.status)
   END_RUNG
   // the same network as SCL:
   "40_UR_R4_DB".DATA.status := "UR1_Robot_status";
END_REGION

REGION Network 2: Copie ETAT UR R5
   RUNG wire#powerrail
      Move(in := "UR2_Robot_status", out1 => "60_UR_R5_DB".DATA.status)
   END_RUNG
   // the same network as SCL:
   "60_UR_R5_DB".DATA.status := "UR2_Robot_status";
END_REGION

REGION Network 3: Copie Registres IN UR R4
   RUNG wire#powerrail
      Move(in := "UR1_Bit_registers", out1 => "40_UR_R4_DB".DATA.Registers.Bit)
      Move(in := "UR1_Int_registers", out1 => "40_UR_R4_DB".DATA.Registers."Int")
      Move(in := "UR1_Float_registers", out1 => "40_UR_R4_DB".DATA.Registers.Float)
   END_RUNG
   // the same network as SCL:
   "40_UR_R4_DB".DATA.Registers.Bit := "UR1_Bit_registers";
   "40_UR_R4_DB".DATA.Registers."Int" := "UR1_Int_registers";
   "40_UR_R4_DB".DATA.Registers.Float := "UR1_Float_registers";
END_REGION

REGION Network 4: Copie Registres IN UR R5
   RUNG wire#powerrail
      Move(in := "UR2_Bit_registers", out1 => "60_UR_R5_DB".DATA.Registers.Bit)
      Move(in := "UR2_Int_registers", out1 => "60_UR_R5_DB".DATA.Registers."Int")
      Move(in := "UR2_Float_registers", out1 => "60_UR_R5_DB".DATA.Registers.Float)
   END_RUNG
   // the same network as SCL:
   "60_UR_R5_DB".DATA.Registers.Bit := "UR2_Bit_registers";
   "60_UR_R5_DB".DATA.Registers."Int" := "UR2_Int_registers";
   "60_UR_R5_DB".DATA.Registers.Float := "UR2_Float_registers";
END_REGION

REGION Network 5: Copie entrees FANUC R1
   RUNG wire#powerrail
      Move(in := "I_FANUC_R1", out1 => "Fanuc_R1_DB".DATA.status)
   END_RUNG
   // the same network as SCL:
   "Fanuc_R1_DB".DATA.status := "I_FANUC_R1";
END_REGION

REGION Network 6: Copie entrees Fanuc R2
   RUNG wire#powerrail
      Move(in := "I_FANUC_R2", out1 => "Fanuc_R2_DB".DATA.status)
   END_RUNG
   // the same network as SCL:
   "Fanuc_R2_DB".DATA.status := "I_FANUC_R2";
END_REGION

REGION Network 7: Copie entrees GoFa R3
   RUNG wire#powerrail
      Move(in := "I_GoFa", out1 => "GoFa_R3_FB_DB".GoFa_Status)
   END_RUNG
   // the same network as SCL:
   "GoFa_R3_FB_DB".GoFa_Status := "I_GoFa";
END_REGION

REGION Network 8: Communication Modbus avec les AGVs
   RUNG wire#powerrail
      "AGVs_Modbus_Read_COM_DB"()
   END_RUNG
   // the same network as SCL:
   "AGVs_Modbus_Read_COM_DB"();   // "AGVs_Modbus_Read_COM"
END_REGION

REGION Network 9: Copie etat Conv01 Conditionnement
   RUNG wire#powerrail
      Move(in := "CV01_Status", out1 => "DB_Variateurs".ConvoyeurC01.Status)
   END_RUNG
   // the same network as SCL:
   "DB_Variateurs".ConvoyeurC01.Status := "CV01_Status";
END_REGION

REGION Network 10: Copie etat Conv02 Conditionnement
   RUNG wire#powerrail
      Move(in := "CV02_Status", out1 => "DB_Variateurs".ConvoyeurC02.Status)
   END_RUNG
   // the same network as SCL:
   "DB_Variateurs".ConvoyeurC02.Status := "CV02_Status";
END_REGION

REGION Network 11: Copie etat Conv03 Conditionnement
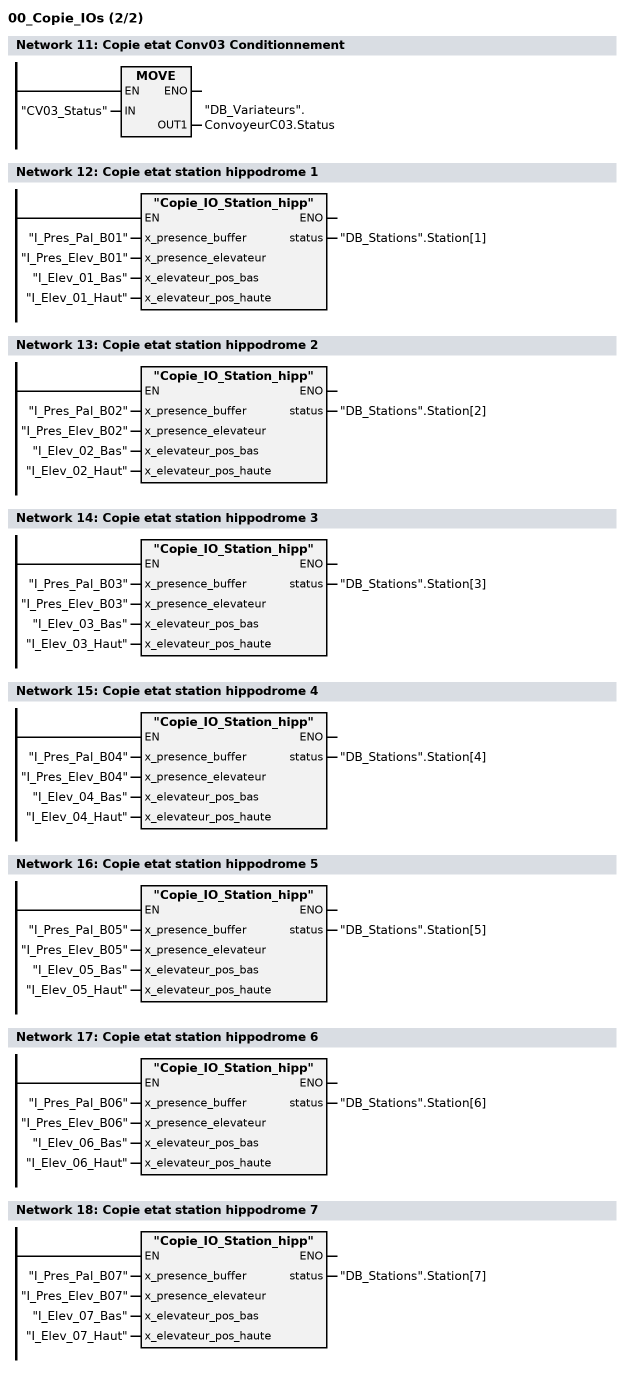
   RUNG wire#powerrail
      Move(in := "CV03_Status", out1 => "DB_Variateurs".ConvoyeurC03.Status)
   END_RUNG
   // the same network as SCL:
   "DB_Variateurs".ConvoyeurC03.Status := "CV03_Status";
END_REGION

REGION Network 12: Copie etat station hippodrome 1
   RUNG wire#powerrail
      "Copie_IO_Station_hipp"(x_presence_buffer := "I_Pres_Pal_B01", x_presence_elevateur := "I_Pres_Elev_B01", x_elevateur_pos_bas := "I_Elev_01_Bas", x_elevateur_pos_haute := "I_Elev_01_Haut", status => "DB_Stations".Station[1])
   END_RUNG
   // the same network as SCL:
   "Copie_IO_Station_hipp"(x_presence_buffer := "I_Pres_Pal_B01",
                           x_presence_elevateur := "I_Pres_Elev_B01",
                           x_elevateur_pos_bas := "I_Elev_01_Bas",
                           x_elevateur_pos_haute := "I_Elev_01_Haut",
                           status => "DB_Stations".Station[1]);
END_REGION

REGION Network 13: Copie etat station hippodrome 2
   RUNG wire#powerrail
      "Copie_IO_Station_hipp"(x_presence_buffer := "I_Pres_Pal_B02", x_presence_elevateur := "I_Pres_Elev_B02", x_elevateur_pos_bas := "I_Elev_02_Bas", x_elevateur_pos_haute := "I_Elev_02_Haut", status => "DB_Stations".Station[2])
   END_RUNG
   // the same network as SCL:
   "Copie_IO_Station_hipp"(x_presence_buffer := "I_Pres_Pal_B02",
                           x_presence_elevateur := "I_Pres_Elev_B02",
                           x_elevateur_pos_bas := "I_Elev_02_Bas",
                           x_elevateur_pos_haute := "I_Elev_02_Haut",
                           status => "DB_Stations".Station[2]);
END_REGION

REGION Network 14: Copie etat station hippodrome 3
   RUNG wire#powerrail
      "Copie_IO_Station_hipp"(x_presence_buffer := "I_Pres_Pal_B03", x_presence_elevateur := "I_Pres_Elev_B03", x_elevateur_pos_bas := "I_Elev_03_Bas", x_elevateur_pos_haute := "I_Elev_03_Haut", status => "DB_Stations".Station[3])
   END_RUNG
   // the same network as SCL:
   "Copie_IO_Station_hipp"(x_presence_buffer := "I_Pres_Pal_B03",
                           x_presence_elevateur := "I_Pres_Elev_B03",
                           x_elevateur_pos_bas := "I_Elev_03_Bas",
                           x_elevateur_pos_haute := "I_Elev_03_Haut",
                           status => "DB_Stations".Station[3]);
END_REGION

REGION Network 15: Copie etat station hippodrome 4
   RUNG wire#powerrail
      "Copie_IO_Station_hipp"(x_presence_buffer := "I_Pres_Pal_B04", x_presence_elevateur := "I_Pres_Elev_B04", x_elevateur_pos_bas := "I_Elev_04_Bas", x_elevateur_pos_haute := "I_Elev_04_Haut", status => "DB_Stations".Station[4])
   END_RUNG
   // the same network as SCL:
   "Copie_IO_Station_hipp"(x_presence_buffer := "I_Pres_Pal_B04",
                           x_presence_elevateur := "I_Pres_Elev_B04",
                           x_elevateur_pos_bas := "I_Elev_04_Bas",
                           x_elevateur_pos_haute := "I_Elev_04_Haut",
                           status => "DB_Stations".Station[4]);
END_REGION

REGION Network 16: Copie etat station hippodrome 5
   RUNG wire#powerrail
      "Copie_IO_Station_hipp"(x_presence_buffer := "I_Pres_Pal_B05", x_presence_elevateur := "I_Pres_Elev_B05", x_elevateur_pos_bas := "I_Elev_05_Bas", x_elevateur_pos_haute := "I_Elev_05_Haut", status => "DB_Stations".Station[5])
   END_RUNG
   // the same network as SCL:
   "Copie_IO_Station_hipp"(x_presence_buffer := "I_Pres_Pal_B05",
                           x_presence_elevateur := "I_Pres_Elev_B05",
                           x_elevateur_pos_bas := "I_Elev_05_Bas",
                           x_elevateur_pos_haute := "I_Elev_05_Haut",
                           status => "DB_Stations".Station[5]);
END_REGION

REGION Network 17: Copie etat station hippodrome 6
   RUNG wire#powerrail
      "Copie_IO_Station_hipp"(x_presence_buffer := "I_Pres_Pal_B06", x_presence_elevateur := "I_Pres_Elev_B06", x_elevateur_pos_bas := "I_Elev_06_Bas", x_elevateur_pos_haute := "I_Elev_06_Haut", status => "DB_Stations".Station[6])
   END_RUNG
   // the same network as SCL:
   "Copie_IO_Station_hipp"(x_presence_buffer := "I_Pres_Pal_B06",
                           x_presence_elevateur := "I_Pres_Elev_B06",
                           x_elevateur_pos_bas := "I_Elev_06_Bas",
                           x_elevateur_pos_haute := "I_Elev_06_Haut",
                           status => "DB_Stations".Station[6]);
END_REGION

REGION Network 18: Copie etat station hippodrome 7
   RUNG wire#powerrail
      "Copie_IO_Station_hipp"(x_presence_buffer := "I_Pres_Pal_B07", x_presence_elevateur := "I_Pres_Elev_B07", x_elevateur_pos_bas := "I_Elev_07_Bas", x_elevateur_pos_haute := "I_Elev_07_Haut", status => "DB_Stations".Station[7])
   END_RUNG
   // the same network as SCL:
   "Copie_IO_Station_hipp"(x_presence_buffer := "I_Pres_Pal_B07",
                           x_presence_elevateur := "I_Pres_Elev_B07",
                           x_elevateur_pos_bas := "I_Elev_07_Bas",
                           x_elevateur_pos_haute := "I_Elev_07_Haut",
                           status => "DB_Stations".Station[7]);
END_REGION
END_FUNCTION

FUNCTION "Copie_IO_Station_hipp" : Void   // FC17, LAD
TITLE = Copie IOs stations hipoddrome
{ S7_Optimized_Access := 'TRUE' }
VERSION : 0.1
   VAR_INPUT
      x_presence_buffer : Bool;
      x_presence_elevateur : Bool;
      x_elevateur_pos_bas : Bool;
      x_elevateur_pos_haute : Bool;
   END_VAR
   VAR_OUTPUT
      status : "Station_Hipp";
   END_VAR
BEGIN

REGION Network 1: Presence palette buffer
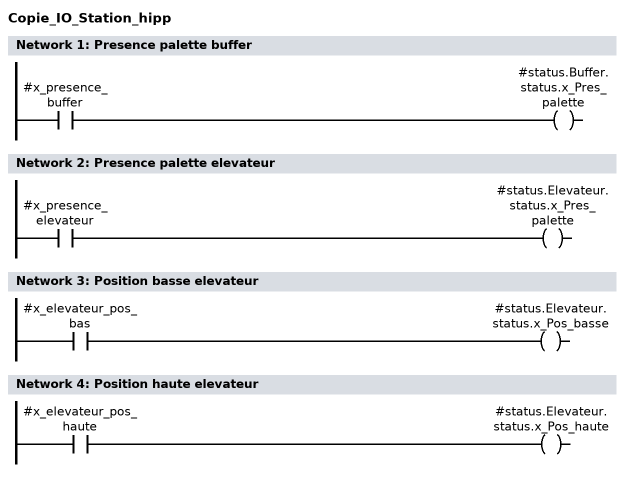
   RUNG wire#powerrail
      Contact( #x_presence_buffer )
      Coil( #status.Buffer.status.x_Pres_palette )
   END_RUNG
   // the same network as SCL:
   #status.Buffer.status.x_Pres_palette := #x_presence_buffer;
END_REGION

REGION Network 2: Presence palette elevateur
   RUNG wire#powerrail
      Contact( #x_presence_elevateur )
      Coil( #status.Elevateur.status.x_Pres_palette )
   END_RUNG
   // the same network as SCL:
   #status.Elevateur.status.x_Pres_palette := #x_presence_elevateur;
END_REGION

REGION Network 3: Position basse elevateur
   RUNG wire#powerrail
      Contact( #x_elevateur_pos_bas )
      Coil( #status.Elevateur.status.x_Pos_basse )
   END_RUNG
   // the same network as SCL:
   #status.Elevateur.status.x_Pos_basse := #x_elevateur_pos_bas;
END_REGION

REGION Network 4: Position haute elevateur
   RUNG wire#powerrail
      Contact( #x_elevateur_pos_haute )
      Coil( #status.Elevateur.status.x_Pos_haute )
   END_RUNG
   // the same network as SCL:
   #status.Elevateur.status.x_Pos_haute := #x_elevateur_pos_haute;
END_REGION
END_FUNCTION

// folder: 100_Gestion_sorties

FUNCTION "101_Gestion_Voyants" : Void   // FC3, LAD
{ S7_Optimized_Access := 'TRUE' }
VERSION : 0.1
BEGIN

REGION Network 1: Voyant HMI Mode Demo
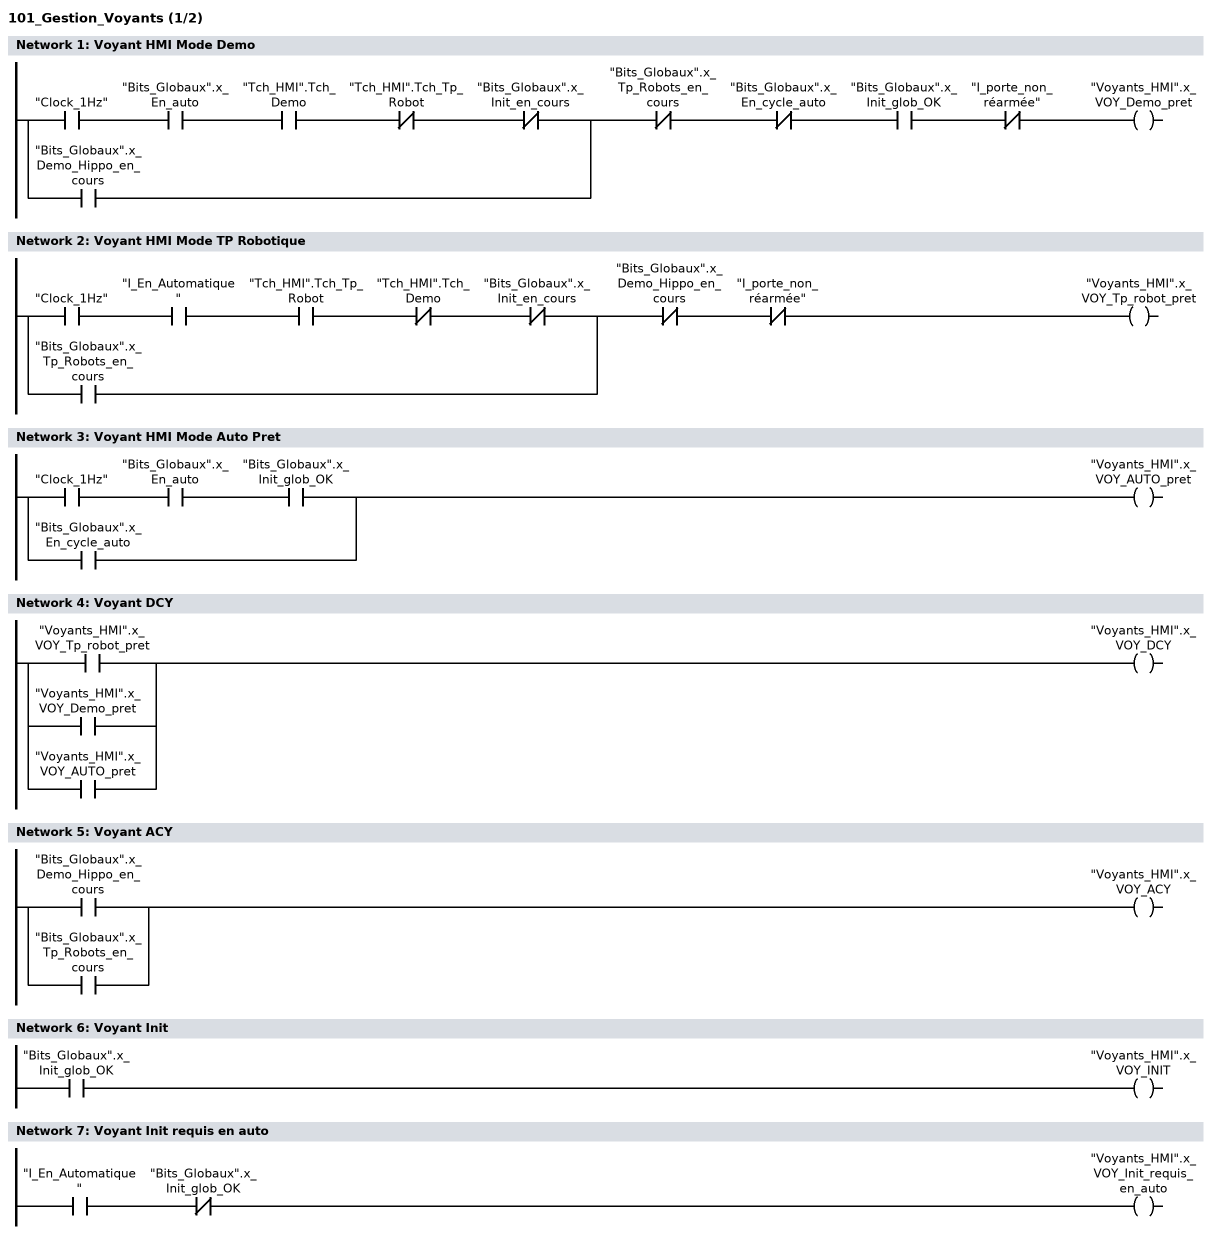
   RUNG wire#powerrail
      Contact( "Clock_1Hz" )
      Contact( "Bits_Globaux".x_En_auto )
      Contact( "Tch_HMI".Tch_Demo )
      I_Contact( "Tch_HMI".Tch_Tp_Robot )
      I_Contact( "Bits_Globaux".x_Init_en_cours )
      wire#w1
      I_Contact( "Bits_Globaux".x_Tp_Robots_en_cours )
      I_Contact( "Bits_Globaux".x_En_cycle_auto )
      Contact( "Bits_Globaux".x_Init_glob_OK )
      I_Contact( "I_porte_non_réarmée" )
      Coil( "Voyants_HMI".x_VOY_Demo_pret )
   END_RUNG
   RUNG wire#powerrail
      Contact( "Bits_Globaux".x_Demo_Hippo_en_cours )
   END_RUNG wire#w1
   // the same network as SCL:
   "Voyants_HMI".x_VOY_Demo_pret := (("Clock_1Hz" AND "Bits_Globaux".x_En_auto AND "Tch_HMI".Tch_Demo AND NOT "Tch_HMI".Tch_Tp_Robot AND NOT "Bits_Globaux".x_Init_en_cours) OR "Bits_Globaux".x_Demo_Hippo_en_cours) AND NOT "Bits_Globaux".x_Tp_Robots_en_cours AND NOT "Bits_Globaux".x_En_cycle_auto AND "Bits_Globaux".x_Init_glob_OK AND NOT "I_porte_non_réarmée";
END_REGION

REGION Network 2: Voyant HMI Mode TP Robotique
   RUNG wire#powerrail
      Contact( "Clock_1Hz" )
      Contact( "I_En_Automatique" )
      Contact( "Tch_HMI".Tch_Tp_Robot )
      I_Contact( "Tch_HMI".Tch_Demo )
      I_Contact( "Bits_Globaux".x_Init_en_cours )
      wire#w1
      I_Contact( "Bits_Globaux".x_Demo_Hippo_en_cours )
      I_Contact( "I_porte_non_réarmée" )
      Coil( "Voyants_HMI".x_VOY_Tp_robot_pret )
   END_RUNG
   RUNG wire#powerrail
      Contact( "Bits_Globaux".x_Tp_Robots_en_cours )
   END_RUNG wire#w1
   // the same network as SCL:
   "Voyants_HMI".x_VOY_Tp_robot_pret := (("Clock_1Hz" AND "I_En_Automatique" AND "Tch_HMI".Tch_Tp_Robot AND NOT "Tch_HMI".Tch_Demo AND NOT "Bits_Globaux".x_Init_en_cours) OR "Bits_Globaux".x_Tp_Robots_en_cours) AND NOT "Bits_Globaux".x_Demo_Hippo_en_cours AND NOT "I_porte_non_réarmée";
END_REGION

REGION Network 3: Voyant HMI Mode Auto Pret
   RUNG wire#powerrail
      Contact( "Clock_1Hz" )
      Contact( "Bits_Globaux".x_En_auto )
      Contact( "Bits_Globaux".x_Init_glob_OK )
      wire#w1
      Coil( "Voyants_HMI".x_VOY_AUTO_pret )
   END_RUNG
   RUNG wire#powerrail
      Contact( "Bits_Globaux".x_En_cycle_auto )
   END_RUNG wire#w1
   // the same network as SCL:
   "Voyants_HMI".x_VOY_AUTO_pret := ("Clock_1Hz" AND "Bits_Globaux".x_En_auto AND "Bits_Globaux".x_Init_glob_OK) OR "Bits_Globaux".x_En_cycle_auto;
END_REGION

REGION Network 4: Voyant DCY
   RUNG wire#powerrail
      Contact( "Voyants_HMI".x_VOY_Tp_robot_pret )
      wire#w1
      Coil( "Voyants_HMI".x_VOY_DCY )
   END_RUNG
   RUNG wire#powerrail
      Contact( "Voyants_HMI".x_VOY_Demo_pret )
   END_RUNG wire#w1
   RUNG wire#powerrail
      Contact( "Voyants_HMI".x_VOY_AUTO_pret )
   END_RUNG wire#w1
   // the same network as SCL:
   "Voyants_HMI".x_VOY_DCY := "Voyants_HMI".x_VOY_Tp_robot_pret OR "Voyants_HMI".x_VOY_Demo_pret OR "Voyants_HMI".x_VOY_AUTO_pret;
END_REGION

REGION Network 5: Voyant ACY
   RUNG wire#powerrail
      Contact( "Bits_Globaux".x_Demo_Hippo_en_cours )
      wire#w1
      Coil( "Voyants_HMI".x_VOY_ACY )
   END_RUNG
   RUNG wire#powerrail
      Contact( "Bits_Globaux".x_Tp_Robots_en_cours )
   END_RUNG wire#w1
   // the same network as SCL:
   "Voyants_HMI".x_VOY_ACY := "Bits_Globaux".x_Demo_Hippo_en_cours OR "Bits_Globaux".x_Tp_Robots_en_cours;
END_REGION

REGION Network 6: Voyant Init
   RUNG wire#powerrail
      Contact( "Bits_Globaux".x_Init_glob_OK )
      Coil( "Voyants_HMI".x_VOY_INIT )
   END_RUNG
   // the same network as SCL:
   "Voyants_HMI".x_VOY_INIT := "Bits_Globaux".x_Init_glob_OK;
END_REGION

REGION Network 7: Voyant Init requis en auto
   RUNG wire#powerrail
      Contact( "I_En_Automatique" )
      I_Contact( "Bits_Globaux".x_Init_glob_OK )
      Coil( "Voyants_HMI".x_VOY_Init_requis_en_auto )
   END_RUNG
   // the same network as SCL:
   "Voyants_HMI".x_VOY_Init_requis_en_auto := "I_En_Automatique" AND NOT "Bits_Globaux".x_Init_glob_OK;
END_REGION

REGION Network 8: Voyant VERT Colonne lumineuse
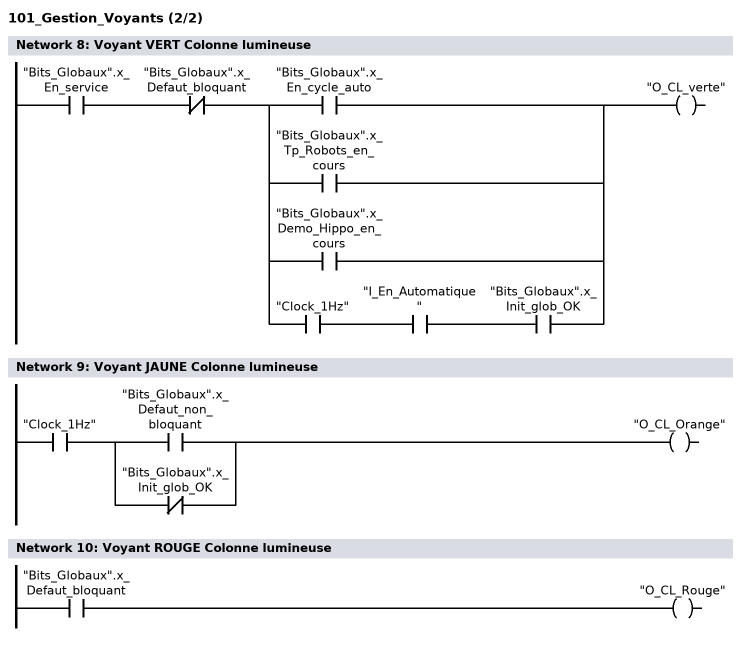
   RUNG wire#powerrail
      Contact( "Bits_Globaux".x_En_service )
      I_Contact( "Bits_Globaux".x_Defaut_bloquant )
      wire#w1
      Contact( "Bits_Globaux".x_En_cycle_auto )
      wire#w2
      Coil( "O_CL_verte" )
   END_RUNG
   RUNG wire#w1
      Contact( "Bits_Globaux".x_Tp_Robots_en_cours )
   END_RUNG wire#w2
   RUNG wire#w1
      Contact( "Bits_Globaux".x_Demo_Hippo_en_cours )
   END_RUNG wire#w2
   RUNG wire#w1
      Contact( "Clock_1Hz" )
      Contact( "I_En_Automatique" )
      Contact( "Bits_Globaux".x_Init_glob_OK )
   END_RUNG wire#w2
   // the same network as SCL:
   "O_CL_verte" := "Bits_Globaux".x_En_service AND NOT "Bits_Globaux".x_Defaut_bloquant AND ("Bits_Globaux".x_En_cycle_auto OR "Bits_Globaux".x_Tp_Robots_en_cours OR "Bits_Globaux".x_Demo_Hippo_en_cours OR ("Clock_1Hz" AND "I_En_Automatique" AND "Bits_Globaux".x_Init_glob_OK));
END_REGION

REGION Network 9: Voyant JAUNE Colonne lumineuse
   RUNG wire#powerrail
      Contact( "Clock_1Hz" )
      wire#w1
      Contact( "Bits_Globaux".x_Defaut_non_bloquant )
      wire#w2
      Coil( "O_CL_Orange" )
   END_RUNG
   RUNG wire#w1
      I_Contact( "Bits_Globaux".x_Init_glob_OK )
   END_RUNG wire#w2
   // the same network as SCL:
   "O_CL_Orange" := "Clock_1Hz" AND ("Bits_Globaux".x_Defaut_non_bloquant OR NOT "Bits_Globaux".x_Init_glob_OK);
END_REGION

REGION Network 10: Voyant ROUGE Colonne lumineuse
   RUNG wire#powerrail
      Contact( "Bits_Globaux".x_Defaut_bloquant )
      Coil( "O_CL_Rouge" )
   END_RUNG
   // the same network as SCL:
   "O_CL_Rouge" := "Bits_Globaux".x_Defaut_bloquant;
END_REGION
END_FUNCTION

FUNCTION "102_Gestion_bits_sortie_virtuels" : Void   // FC5, LAD
{ S7_Optimized_Access := 'TRUE' }
VERSION : 0.1
BEGIN

REGION Network 1: Confirmation cobots et Robots en auto
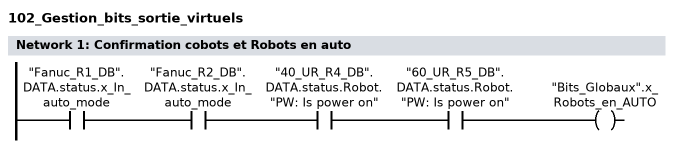
   RUNG wire#powerrail
      Contact( "Fanuc_R1_DB".DATA.status.x_In_auto_mode )
      Contact( "Fanuc_R2_DB".DATA.status.x_In_auto_mode )
      Contact( "40_UR_R4_DB".DATA.status.Robot."PW: Is power on" )
      Contact( "60_UR_R5_DB".DATA.status.Robot."PW: Is power on" )
      Coil( "Bits_Globaux".x_Robots_en_AUTO )
   END_RUNG
   // the same network as SCL:
   "Bits_Globaux".x_Robots_en_AUTO := "Fanuc_R1_DB".DATA.status.x_In_auto_mode AND "Fanuc_R2_DB".DATA.status.x_In_auto_mode AND "40_UR_R4_DB".DATA.status.Robot."PW: Is power on" AND "60_UR_R5_DB".DATA.status.Robot."PW: Is power on";
END_REGION
END_FUNCTION

FUNCTION "103_Gestion_Bits_Imprimantes" : Void   // FC7, LAD
{ S7_Optimized_Access := 'TRUE' }
VERSION : 0.1
BEGIN
END_FUNCTION

FUNCTION "104_Gestion_Bits_Keyence" : Void   // FC8, LAD
{ S7_Optimized_Access := 'TRUE' }
VERSION : 0.1
BEGIN
END_FUNCTION

FUNCTION "105_Gestion_Bits_Cobots" : Void   // FC10, LAD
{ S7_Optimized_Access := 'TRUE' }
VERSION : 0.1
BEGIN

REGION Network 1: Cobot UR4
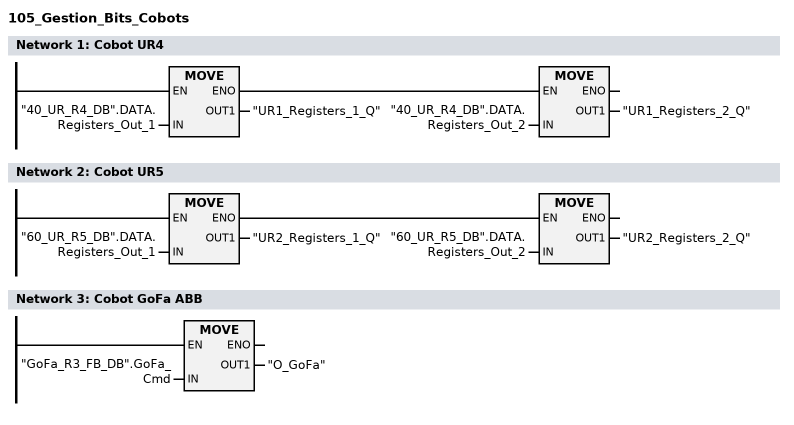
   RUNG wire#powerrail
      Move(in := "40_UR_R4_DB".DATA.Registers_Out_1, out1 => "UR1_Registers_1_Q")
      Move(in := "40_UR_R4_DB".DATA.Registers_Out_2, out1 => "UR1_Registers_2_Q")
   END_RUNG
   // the same network as SCL:
   "UR1_Registers_1_Q" := "40_UR_R4_DB".DATA.Registers_Out_1;
   "UR1_Registers_2_Q" := "40_UR_R4_DB".DATA.Registers_Out_2;
END_REGION

REGION Network 2: Cobot UR5
   RUNG wire#powerrail
      Move(in := "60_UR_R5_DB".DATA.Registers_Out_1, out1 => "UR2_Registers_1_Q")
      Move(in := "60_UR_R5_DB".DATA.Registers_Out_2, out1 => "UR2_Registers_2_Q")
   END_RUNG
   // the same network as SCL:
   "UR2_Registers_1_Q" := "60_UR_R5_DB".DATA.Registers_Out_1;
   "UR2_Registers_2_Q" := "60_UR_R5_DB".DATA.Registers_Out_2;
END_REGION

REGION Network 3: Cobot GoFa ABB
   RUNG wire#powerrail
      Move(in := "GoFa_R3_FB_DB".GoFa_Cmd, out1 => "O_GoFa")
   END_RUNG
   // the same network as SCL:
   "O_GoFa" := "GoFa_R3_FB_DB".GoFa_Cmd;
END_REGION
END_FUNCTION

FUNCTION "106_Gestion_Bits_Robots" : Void   // FC11, LAD
{ S7_Optimized_Access := 'TRUE' }
VERSION : 0.1
BEGIN

REGION Network 1: Fanuc R1 Sorties
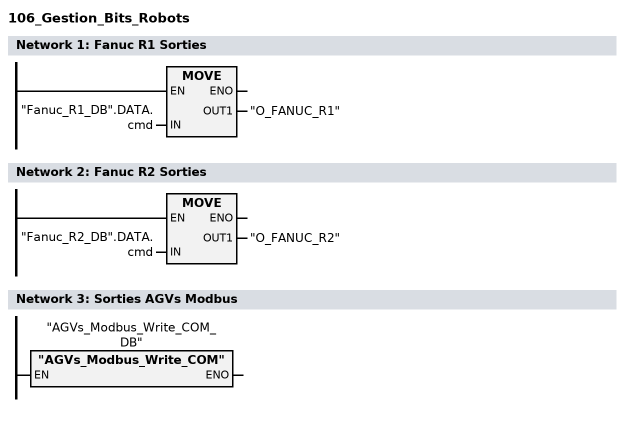
   RUNG wire#powerrail
      Move(in := "Fanuc_R1_DB".DATA.cmd, out1 => "O_FANUC_R1")
   END_RUNG
   // the same network as SCL:
   "O_FANUC_R1" := "Fanuc_R1_DB".DATA.cmd;
END_REGION

REGION Network 2: Fanuc R2 Sorties
   RUNG wire#powerrail
      Move(in := "Fanuc_R2_DB".DATA.cmd, out1 => "O_FANUC_R2")
   END_RUNG
   // the same network as SCL:
   "O_FANUC_R2" := "Fanuc_R2_DB".DATA.cmd;
END_REGION

REGION Network 3: Sorties AGVs Modbus
   RUNG wire#powerrail
      "AGVs_Modbus_Write_COM_DB"()
   END_RUNG
   // the same network as SCL:
   "AGVs_Modbus_Write_COM_DB"();   // "AGVs_Modbus_Write_COM"
END_REGION
END_FUNCTION

FUNCTION "107_Gestion_des_portes" : Void   // FC12, LAD
TITLE = Gestion des portes d'acces
{ S7_Optimized_Access := 'TRUE' }
VERSION : 0.1
BEGIN

REGION Network 1: Autorisation ouverture porte
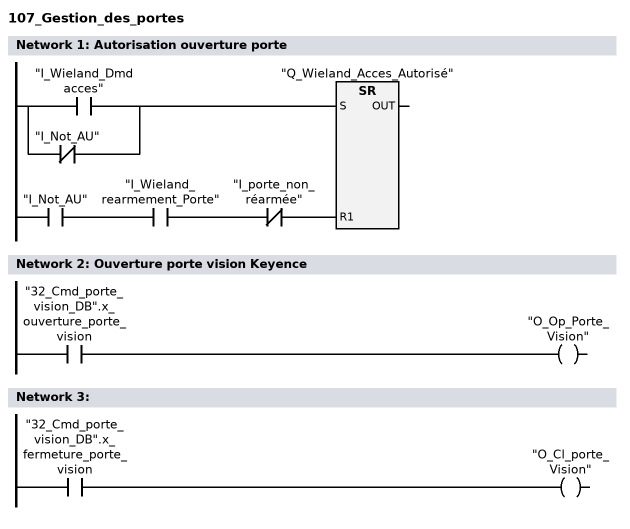
   RUNG wire#powerrail
      Contact( "I_Wieland_Dmd acces" )
      wire#w1
      S_SR(operand := "Q_Wieland_Acces_Autorisé", r1 := wire#w2)
   END_RUNG
   RUNG wire#powerrail
      I_Contact( "I_Not_AU" )
   END_RUNG wire#w1
   RUNG wire#powerrail
      Contact( "I_Not_AU" )
      Contact( "I_Wieland_rearmement_Porte" )
      I_Contact( "I_porte_non_réarmée" )
   END_RUNG wire#w2
   // the same network as SCL:
   IF "I_Wieland_Dmd acces" OR NOT "I_Not_AU" THEN
       "Q_Wieland_Acces_Autorisé" := TRUE;   // SR flip-flop
   END_IF;
   IF "I_Not_AU" AND "I_Wieland_rearmement_Porte" AND NOT "I_porte_non_réarmée" THEN
       "Q_Wieland_Acces_Autorisé" := FALSE;
   END_IF;
END_REGION

REGION Network 2: Ouverture porte vision Keyence
   RUNG wire#powerrail
      Contact( "32_Cmd_porte_vision_DB".x_ouverture_porte_vision )
      Coil( "O_Op_Porte_Vision" )
   END_RUNG
   // the same network as SCL:
   "O_Op_Porte_Vision" := "32_Cmd_porte_vision_DB".x_ouverture_porte_vision;
END_REGION

REGION Network 3
   RUNG wire#powerrail
      Contact( "32_Cmd_porte_vision_DB".x_fermeture_porte_vision )
      Coil( "O_Cl_porte_Vision" )
   END_RUNG
   // the same network as SCL:
   "O_Cl_porte_Vision" := "32_Cmd_porte_vision_DB".x_fermeture_porte_vision;
END_REGION
END_FUNCTION

FUNCTION "108_Gestion_sorties_variateurs" : Void   // FC14, LAD
TITLE = Gestion sortie des variateurs
{ S7_Optimized_Access := 'TRUE' }
VERSION : 0.1
BEGIN

REGION Network 1: Envoi cmd VAR1 (de gauche à droite dans l'armoire)
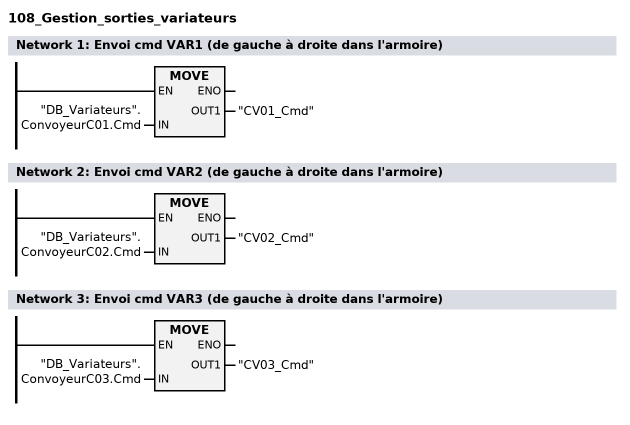
   RUNG wire#powerrail
      Move(in := "DB_Variateurs".ConvoyeurC01.Cmd, out1 => "CV01_Cmd")
   END_RUNG
   // the same network as SCL:
   "CV01_Cmd" := "DB_Variateurs".ConvoyeurC01.Cmd;
END_REGION

REGION Network 2: Envoi cmd VAR2 (de gauche à droite dans l'armoire)
   RUNG wire#powerrail
      Move(in := "DB_Variateurs".ConvoyeurC02.Cmd, out1 => "CV02_Cmd")
   END_RUNG
   // the same network as SCL:
   "CV02_Cmd" := "DB_Variateurs".ConvoyeurC02.Cmd;
END_REGION

REGION Network 3: Envoi cmd VAR3 (de gauche à droite dans l'armoire)
   RUNG wire#powerrail
      Move(in := "DB_Variateurs".ConvoyeurC03.Cmd, out1 => "CV03_Cmd")
   END_RUNG
   // the same network as SCL:
   "CV03_Cmd" := "DB_Variateurs".ConvoyeurC03.Cmd;
END_REGION
END_FUNCTION

FUNCTION "109-Gestion_sorties_conv_hippodrome" : Void   // FC15, LAD
TITLE = Gestion sorties convoyeur hippodrome
{ S7_Optimized_Access := 'TRUE' }
VERSION : 0.1
BEGIN

REGION Network 1: Conv1
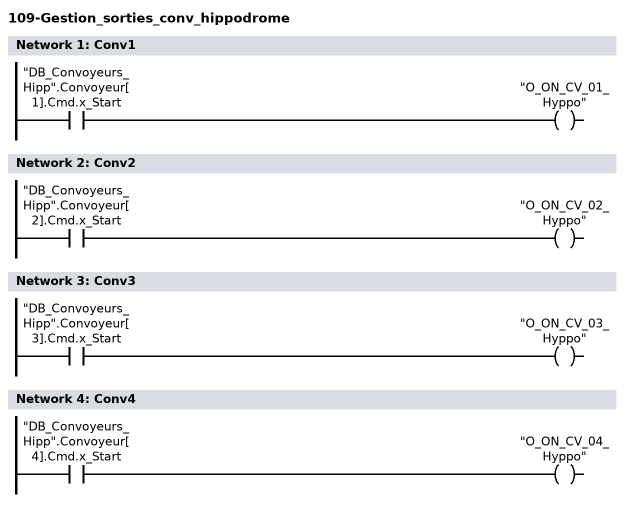
   RUNG wire#powerrail
      Contact( "DB_Convoyeurs_Hipp".Convoyeur[1].Cmd.x_Start )
      Coil( "O_ON_CV_01_Hyppo" )
   END_RUNG
   // the same network as SCL:
   "O_ON_CV_01_Hyppo" := "DB_Convoyeurs_Hipp".Convoyeur[1].Cmd.x_Start;
END_REGION

REGION Network 2: Conv2
   RUNG wire#powerrail
      Contact( "DB_Convoyeurs_Hipp".Convoyeur[2].Cmd.x_Start )
      Coil( "O_ON_CV_02_Hyppo" )
   END_RUNG
   // the same network as SCL:
   "O_ON_CV_02_Hyppo" := "DB_Convoyeurs_Hipp".Convoyeur[2].Cmd.x_Start;
END_REGION

REGION Network 3: Conv3
   RUNG wire#powerrail
      Contact( "DB_Convoyeurs_Hipp".Convoyeur[3].Cmd.x_Start )
      Coil( "O_ON_CV_03_Hyppo" )
   END_RUNG
   // the same network as SCL:
   "O_ON_CV_03_Hyppo" := "DB_Convoyeurs_Hipp".Convoyeur[3].Cmd.x_Start;
END_REGION

REGION Network 4: Conv4
   RUNG wire#powerrail
      Contact( "DB_Convoyeurs_Hipp".Convoyeur[4].Cmd.x_Start )
      Coil( "O_ON_CV_04_Hyppo" )
   END_RUNG
   // the same network as SCL:
   "O_ON_CV_04_Hyppo" := "DB_Convoyeurs_Hipp".Convoyeur[4].Cmd.x_Start;
END_REGION
END_FUNCTION

FUNCTION "110_Gestion_sorties_postes_de_travail" : Void   // FC18, LAD
{ S7_Optimized_Access := 'TRUE' }
VERSION : 0.1
BEGIN

REGION Network 1: CMD poste de travail Hippodrome 1
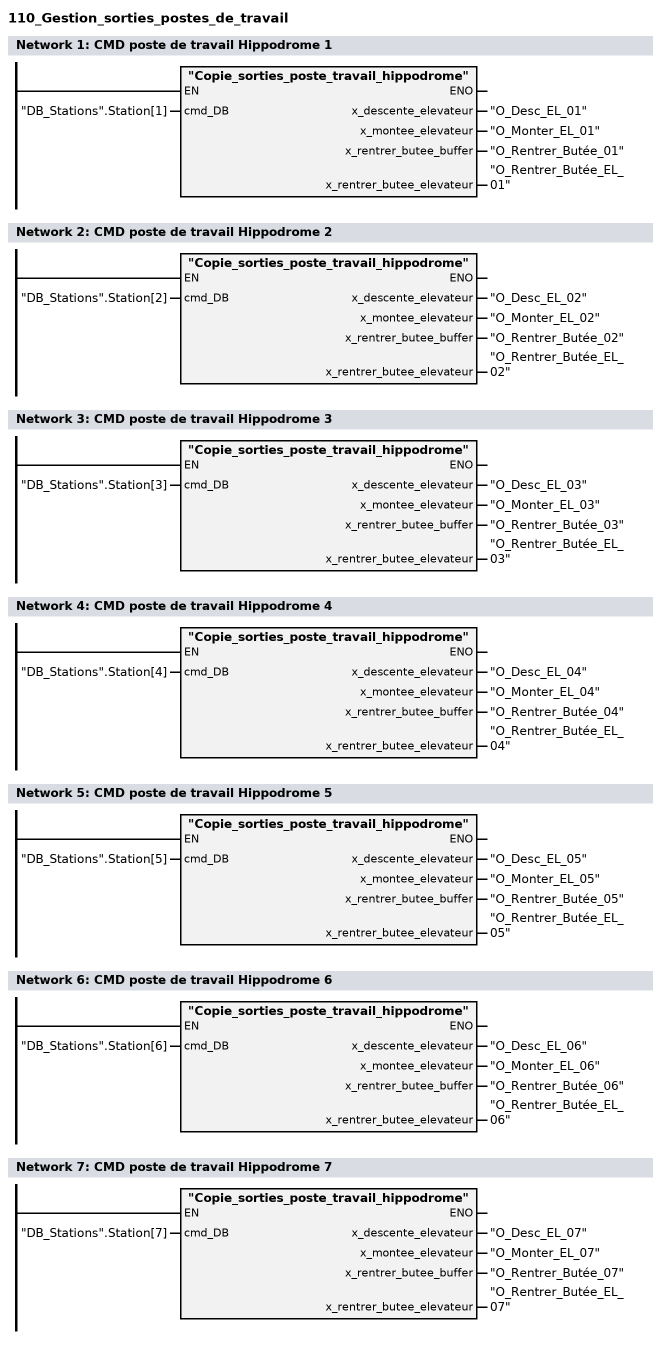
   RUNG wire#powerrail
      "Copie_sorties_poste_travail_hippodrome"(cmd_DB := "DB_Stations".Station[1], x_descente_elevateur => "O_Desc_EL_01", x_montee_elevateur => "O_Monter_EL_01", x_rentrer_butee_buffer => "O_Rentrer_Butée_01", x_rentrer_butee_elevateur => "O_Rentrer_Butée_EL_01")
   END_RUNG
   // the same network as SCL:
   "Copie_sorties_poste_travail_hippodrome"(cmd_DB := "DB_Stations".Station[1],
                           x_descente_elevateur => "O_Desc_EL_01",
                           x_montee_elevateur => "O_Monter_EL_01",
                           x_rentrer_butee_buffer => "O_Rentrer_Butée_01",
                           x_rentrer_butee_elevateur => "O_Rentrer_Butée_EL_01");
END_REGION

REGION Network 2: CMD poste de travail Hippodrome 2
   RUNG wire#powerrail
      "Copie_sorties_poste_travail_hippodrome"(cmd_DB := "DB_Stations".Station[2], x_descente_elevateur => "O_Desc_EL_02", x_montee_elevateur => "O_Monter_EL_02", x_rentrer_butee_buffer => "O_Rentrer_Butée_02", x_rentrer_butee_elevateur => "O_Rentrer_Butée_EL_02")
   END_RUNG
   // the same network as SCL:
   "Copie_sorties_poste_travail_hippodrome"(cmd_DB := "DB_Stations".Station[2],
                           x_descente_elevateur => "O_Desc_EL_02",
                           x_montee_elevateur => "O_Monter_EL_02",
                           x_rentrer_butee_buffer => "O_Rentrer_Butée_02",
                           x_rentrer_butee_elevateur => "O_Rentrer_Butée_EL_02");
END_REGION

REGION Network 3: CMD poste de travail Hippodrome 3
   RUNG wire#powerrail
      "Copie_sorties_poste_travail_hippodrome"(cmd_DB := "DB_Stations".Station[3], x_descente_elevateur => "O_Desc_EL_03", x_montee_elevateur => "O_Monter_EL_03", x_rentrer_butee_buffer => "O_Rentrer_Butée_03", x_rentrer_butee_elevateur => "O_Rentrer_Butée_EL_03")
   END_RUNG
   // the same network as SCL:
   "Copie_sorties_poste_travail_hippodrome"(cmd_DB := "DB_Stations".Station[3],
                           x_descente_elevateur => "O_Desc_EL_03",
                           x_montee_elevateur => "O_Monter_EL_03",
                           x_rentrer_butee_buffer => "O_Rentrer_Butée_03",
                           x_rentrer_butee_elevateur => "O_Rentrer_Butée_EL_03");
END_REGION

REGION Network 4: CMD poste de travail Hippodrome 4
   RUNG wire#powerrail
      "Copie_sorties_poste_travail_hippodrome"(cmd_DB := "DB_Stations".Station[4], x_descente_elevateur => "O_Desc_EL_04", x_montee_elevateur => "O_Monter_EL_04", x_rentrer_butee_buffer => "O_Rentrer_Butée_04", x_rentrer_butee_elevateur => "O_Rentrer_Butée_EL_04")
   END_RUNG
   // the same network as SCL:
   "Copie_sorties_poste_travail_hippodrome"(cmd_DB := "DB_Stations".Station[4],
                           x_descente_elevateur => "O_Desc_EL_04",
                           x_montee_elevateur => "O_Monter_EL_04",
                           x_rentrer_butee_buffer => "O_Rentrer_Butée_04",
                           x_rentrer_butee_elevateur => "O_Rentrer_Butée_EL_04");
END_REGION

REGION Network 5: CMD poste de travail Hippodrome 5
   RUNG wire#powerrail
      "Copie_sorties_poste_travail_hippodrome"(cmd_DB := "DB_Stations".Station[5], x_descente_elevateur => "O_Desc_EL_05", x_montee_elevateur => "O_Monter_EL_05", x_rentrer_butee_buffer => "O_Rentrer_Butée_05", x_rentrer_butee_elevateur => "O_Rentrer_Butée_EL_05")
   END_RUNG
   // the same network as SCL:
   "Copie_sorties_poste_travail_hippodrome"(cmd_DB := "DB_Stations".Station[5],
                           x_descente_elevateur => "O_Desc_EL_05",
                           x_montee_elevateur => "O_Monter_EL_05",
                           x_rentrer_butee_buffer => "O_Rentrer_Butée_05",
                           x_rentrer_butee_elevateur => "O_Rentrer_Butée_EL_05");
END_REGION

REGION Network 6: CMD poste de travail Hippodrome 6
   RUNG wire#powerrail
      "Copie_sorties_poste_travail_hippodrome"(cmd_DB := "DB_Stations".Station[6], x_descente_elevateur => "O_Desc_EL_06", x_montee_elevateur => "O_Monter_EL_06", x_rentrer_butee_buffer => "O_Rentrer_Butée_06", x_rentrer_butee_elevateur => "O_Rentrer_Butée_EL_06")
   END_RUNG
   // the same network as SCL:
   "Copie_sorties_poste_travail_hippodrome"(cmd_DB := "DB_Stations".Station[6],
                           x_descente_elevateur => "O_Desc_EL_06",
                           x_montee_elevateur => "O_Monter_EL_06",
                           x_rentrer_butee_buffer => "O_Rentrer_Butée_06",
                           x_rentrer_butee_elevateur => "O_Rentrer_Butée_EL_06");
END_REGION

REGION Network 7: CMD poste de travail Hippodrome 7
   RUNG wire#powerrail
      "Copie_sorties_poste_travail_hippodrome"(cmd_DB := "DB_Stations".Station[7], x_descente_elevateur => "O_Desc_EL_07", x_montee_elevateur => "O_Monter_EL_07", x_rentrer_butee_buffer => "O_Rentrer_Butée_07", x_rentrer_butee_elevateur => "O_Rentrer_Butée_EL_07")
   END_RUNG
   // the same network as SCL:
   "Copie_sorties_poste_travail_hippodrome"(cmd_DB := "DB_Stations".Station[7],
                           x_descente_elevateur => "O_Desc_EL_07",
                           x_montee_elevateur => "O_Monter_EL_07",
                           x_rentrer_butee_buffer => "O_Rentrer_Butée_07",
                           x_rentrer_butee_elevateur => "O_Rentrer_Butée_EL_07");
END_REGION
END_FUNCTION

FUNCTION "Copie_sorties_poste_travail_hippodrome" : Void   // FC19, LAD
TITLE = Envoi bits de cmd poste de travail hippodrome
{ S7_Optimized_Access := 'TRUE' }
VERSION : 0.1
   VAR_INPUT
      cmd_DB : "Station_Hipp";
   END_VAR
   VAR_OUTPUT
      x_descente_elevateur : Bool;
      x_montee_elevateur : Bool;
      x_rentrer_butee_buffer : Bool;
      x_rentrer_butee_elevateur : Bool;
   END_VAR
BEGIN

REGION Network 1: Descente elevateur
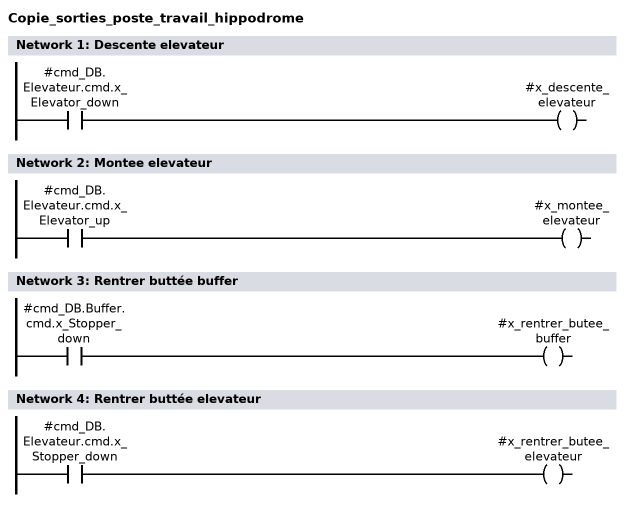
   RUNG wire#powerrail
      Contact( #cmd_DB.Elevateur.cmd.x_Elevator_down )
      Coil( #x_descente_elevateur )
   END_RUNG
   // the same network as SCL:
   #x_descente_elevateur := #cmd_DB.Elevateur.cmd.x_Elevator_down;
END_REGION

REGION Network 2: Montee elevateur
   RUNG wire#powerrail
      Contact( #cmd_DB.Elevateur.cmd.x_Elevator_up )
      Coil( #x_montee_elevateur )
   END_RUNG
   // the same network as SCL:
   #x_montee_elevateur := #cmd_DB.Elevateur.cmd.x_Elevator_up;
END_REGION

REGION Network 3: Rentrer buttée buffer
   RUNG wire#powerrail
      Contact( #cmd_DB.Buffer.cmd.x_Stopper_down )
      Coil( #x_rentrer_butee_buffer )
   END_RUNG
   // the same network as SCL:
   #x_rentrer_butee_buffer := #cmd_DB.Buffer.cmd.x_Stopper_down;
END_REGION

REGION Network 4: Rentrer buttée elevateur
   RUNG wire#powerrail
      Contact( #cmd_DB.Elevateur.cmd.x_Stopper_down )
      Coil( #x_rentrer_butee_elevateur )
   END_RUNG
   // the same network as SCL:
   #x_rentrer_butee_elevateur := #cmd_DB.Elevateur.cmd.x_Stopper_down;
END_REGION
END_FUNCTION

FUNCTION "100_Gestion_sorties" : Void   // FC100, LAD
{ S7_Optimized_Access := 'TRUE' }
VERSION : 0.1
BEGIN

REGION Network 1: Gestion des voyants
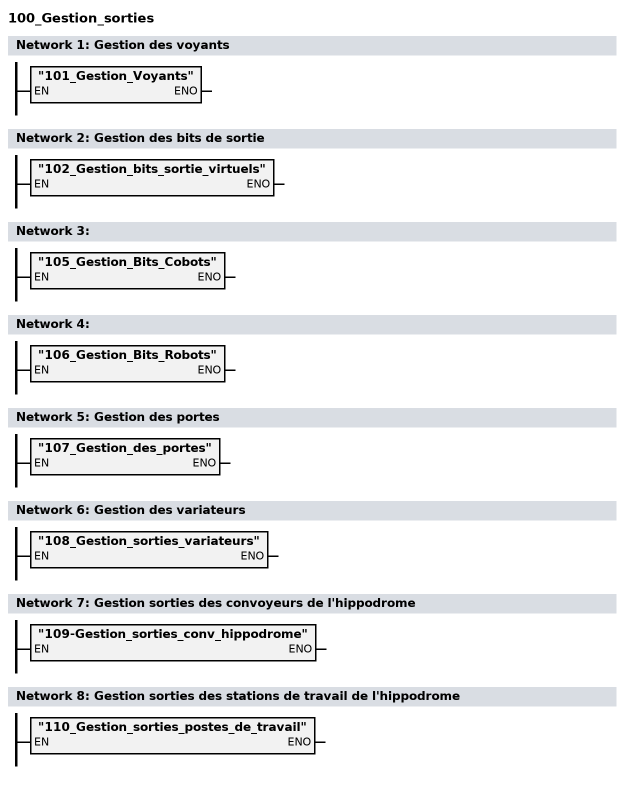
   RUNG wire#powerrail
      "101_Gestion_Voyants"()
   END_RUNG
   // the same network as SCL:
   "101_Gestion_Voyants"();
END_REGION

REGION Network 2: Gestion des bits de sortie
   RUNG wire#powerrail
      "102_Gestion_bits_sortie_virtuels"()
   END_RUNG
   // the same network as SCL:
   "102_Gestion_bits_sortie_virtuels"();
END_REGION

REGION Network 3
   RUNG wire#powerrail
      "105_Gestion_Bits_Cobots"()
   END_RUNG
   // the same network as SCL:
   "105_Gestion_Bits_Cobots"();
END_REGION

REGION Network 4
   RUNG wire#powerrail
      "106_Gestion_Bits_Robots"()
   END_RUNG
   // the same network as SCL:
   "106_Gestion_Bits_Robots"();
END_REGION

REGION Network 5: Gestion des portes
   RUNG wire#powerrail
      "107_Gestion_des_portes"()
   END_RUNG
   // the same network as SCL:
   "107_Gestion_des_portes"();
END_REGION

REGION Network 6: Gestion des variateurs
   RUNG wire#powerrail
      "108_Gestion_sorties_variateurs"()
   END_RUNG
   // the same network as SCL:
   "108_Gestion_sorties_variateurs"();
END_REGION

REGION Network 7: Gestion sorties des convoyeurs de l'hippodrome
   RUNG wire#powerrail
      "109-Gestion_sorties_conv_hippodrome"()
   END_RUNG
   // the same network as SCL:
   "109-Gestion_sorties_conv_hippodrome"();
END_REGION

REGION Network 8: Gestion sorties des stations de travail de l'hippodrome
   RUNG wire#powerrail
      "110_Gestion_sorties_postes_de_travail"()
   END_RUNG
   // the same network as SCL:
   "110_Gestion_sorties_postes_de_travail"();
END_REGION
END_FUNCTION

// folder: 1_Imprimantes_3D

FUNCTION "20_Imprimantes_3D" : Void   // FC2, LAD
{ S7_Optimized_Access := 'TRUE' }
VERSION : 0.1
BEGIN
END_FUNCTION

// folder: 2-Hippodrome

FUNCTION "20-Gestion_equipement_hippodrome" : Void   // FC4, LAD
TITLE = Gestion equipement hippodrome
{ S7_Optimized_Access := 'TRUE' }
VERSION : 0.1
BEGIN

REGION Network 1: Gestion des convoyeurs
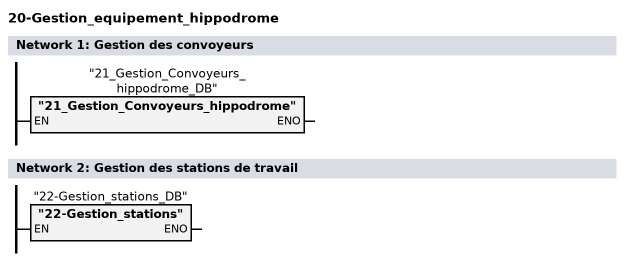
   RUNG wire#powerrail
      "21_Gestion_Convoyeurs_hippodrome_DB"()
   END_RUNG
   // the same network as SCL:
   "21_Gestion_Convoyeurs_hippodrome_DB"();   // "21_Gestion_Convoyeurs_hippodrome"
END_REGION

REGION Network 2: Gestion des stations de travail
   RUNG wire#powerrail
      "22-Gestion_stations_DB"()
   END_RUNG
   // the same network as SCL:
   "22-Gestion_stations_DB"();   // "22-Gestion_stations"
END_REGION
END_FUNCTION

// folder: 2-Hippodrome/Convoyeurs

FUNCTION_BLOCK "Convoyeur_Hippodrome"   // FB8, LAD
TITLE = Pilotage Convoyeur hippodrome
{ S7_Optimized_Access := 'TRUE' }
VERSION : 0.1
   VAR_INPUT
      x_Defaut_externe : Bool;
      x_enService : Bool;
      x_Marche_auto : Bool;
      x_Marche_manu : Bool;
      x_Arret_auto : Bool;
      x_Arret_Manu : Bool;
      x_Retour_defaut_thermique : Bool;
   END_VAR
   VAR_OUTPUT
      Defaut : Bool;
   END_VAR
   VAR_IN_OUT
      DB_Convoyeur_DATA : "Convoyeur_Hipp";
   END_VAR
BEGIN

REGION Network 1: Vérification défaut thermique
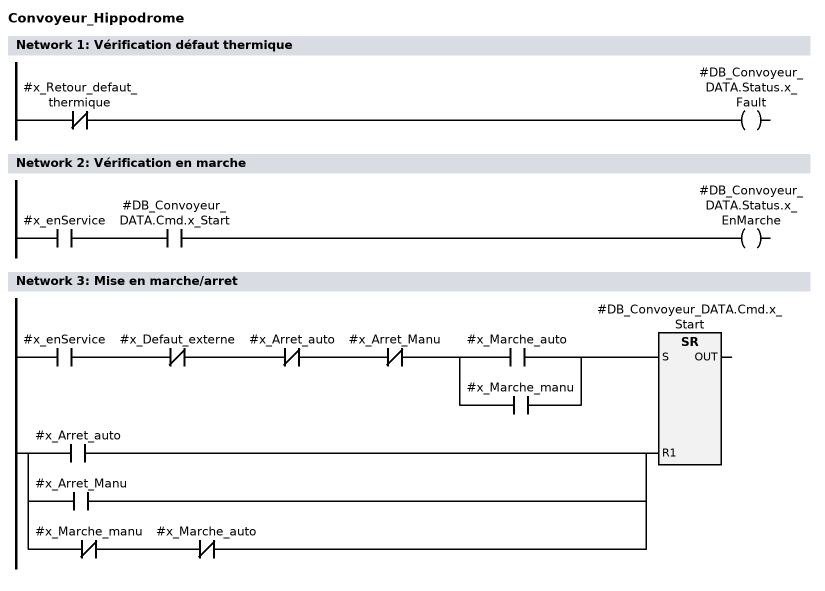
   RUNG wire#powerrail
      I_Contact( #x_Retour_defaut_thermique )
      Coil( #DB_Convoyeur_DATA.Status.x_Fault )
   END_RUNG
   // the same network as SCL:
   #DB_Convoyeur_DATA.Status.x_Fault := NOT #x_Retour_defaut_thermique;
END_REGION

REGION Network 2: Vérification en marche
   RUNG wire#powerrail
      Contact( #x_enService )
      Contact( #DB_Convoyeur_DATA.Cmd.x_Start )
      Coil( #DB_Convoyeur_DATA.Status.x_EnMarche )
   END_RUNG
   // the same network as SCL:
   #DB_Convoyeur_DATA.Status.x_EnMarche := #x_enService AND #DB_Convoyeur_DATA.Cmd.x_Start;
END_REGION

REGION Network 3: Mise en marche/arret
   RUNG wire#powerrail
      Contact( #x_enService )
      I_Contact( #x_Defaut_externe )
      I_Contact( #x_Arret_auto )
      I_Contact( #x_Arret_Manu )
      wire#w1
      Contact( #x_Marche_auto )
      wire#w2
      S_SR(operand := #DB_Convoyeur_DATA.Cmd.x_Start, r1 := wire#w3)
   END_RUNG
   RUNG wire#w1
      Contact( #x_Marche_manu )
   END_RUNG wire#w2
   RUNG wire#powerrail
      Contact( #x_Arret_auto )
   END_RUNG wire#w3
   RUNG wire#powerrail
      Contact( #x_Arret_Manu )
   END_RUNG wire#w3
   RUNG wire#powerrail
      I_Contact( #x_Marche_manu )
      I_Contact( #x_Marche_auto )
   END_RUNG wire#w3
   // the same network as SCL:
   IF #x_enService AND NOT #x_Defaut_externe AND NOT #x_Arret_auto AND NOT #x_Arret_Manu AND (#x_Marche_auto OR #x_Marche_manu) THEN
       #DB_Convoyeur_DATA.Cmd.x_Start := TRUE;   // SR flip-flop
   END_IF;
   IF #x_Arret_auto OR #x_Arret_Manu OR (NOT #x_Marche_manu AND NOT #x_Marche_auto) THEN
       #DB_Convoyeur_DATA.Cmd.x_Start := FALSE;
   END_IF;
END_REGION
END_FUNCTION_BLOCK

FUNCTION_BLOCK "21_Gestion_Convoyeurs_hippodrome"   // FB9, LAD
TITLE = Gestion des convoyeurs de l'hippodrome
{ S7_Optimized_Access := 'TRUE' }
VERSION : 0.1
   VAR
      Convoyeur_Hippodrome_1 : "Convoyeur_Hippodrome";
      Convoyeur_Hippodrome_2 : "Convoyeur_Hippodrome";
      Convoyeur_Hippodrome_3 : "Convoyeur_Hippodrome";
      Convoyeur_Hippodrome_4 : "Convoyeur_Hippodrome";
      x_All_stations_empty : Bool;
      Timer_attente_arret_convoyeurs : TON_TIME;
   END_VAR
BEGIN

REGION Network 1: Arret convoyeurs en auto si toutes les stations sont vides
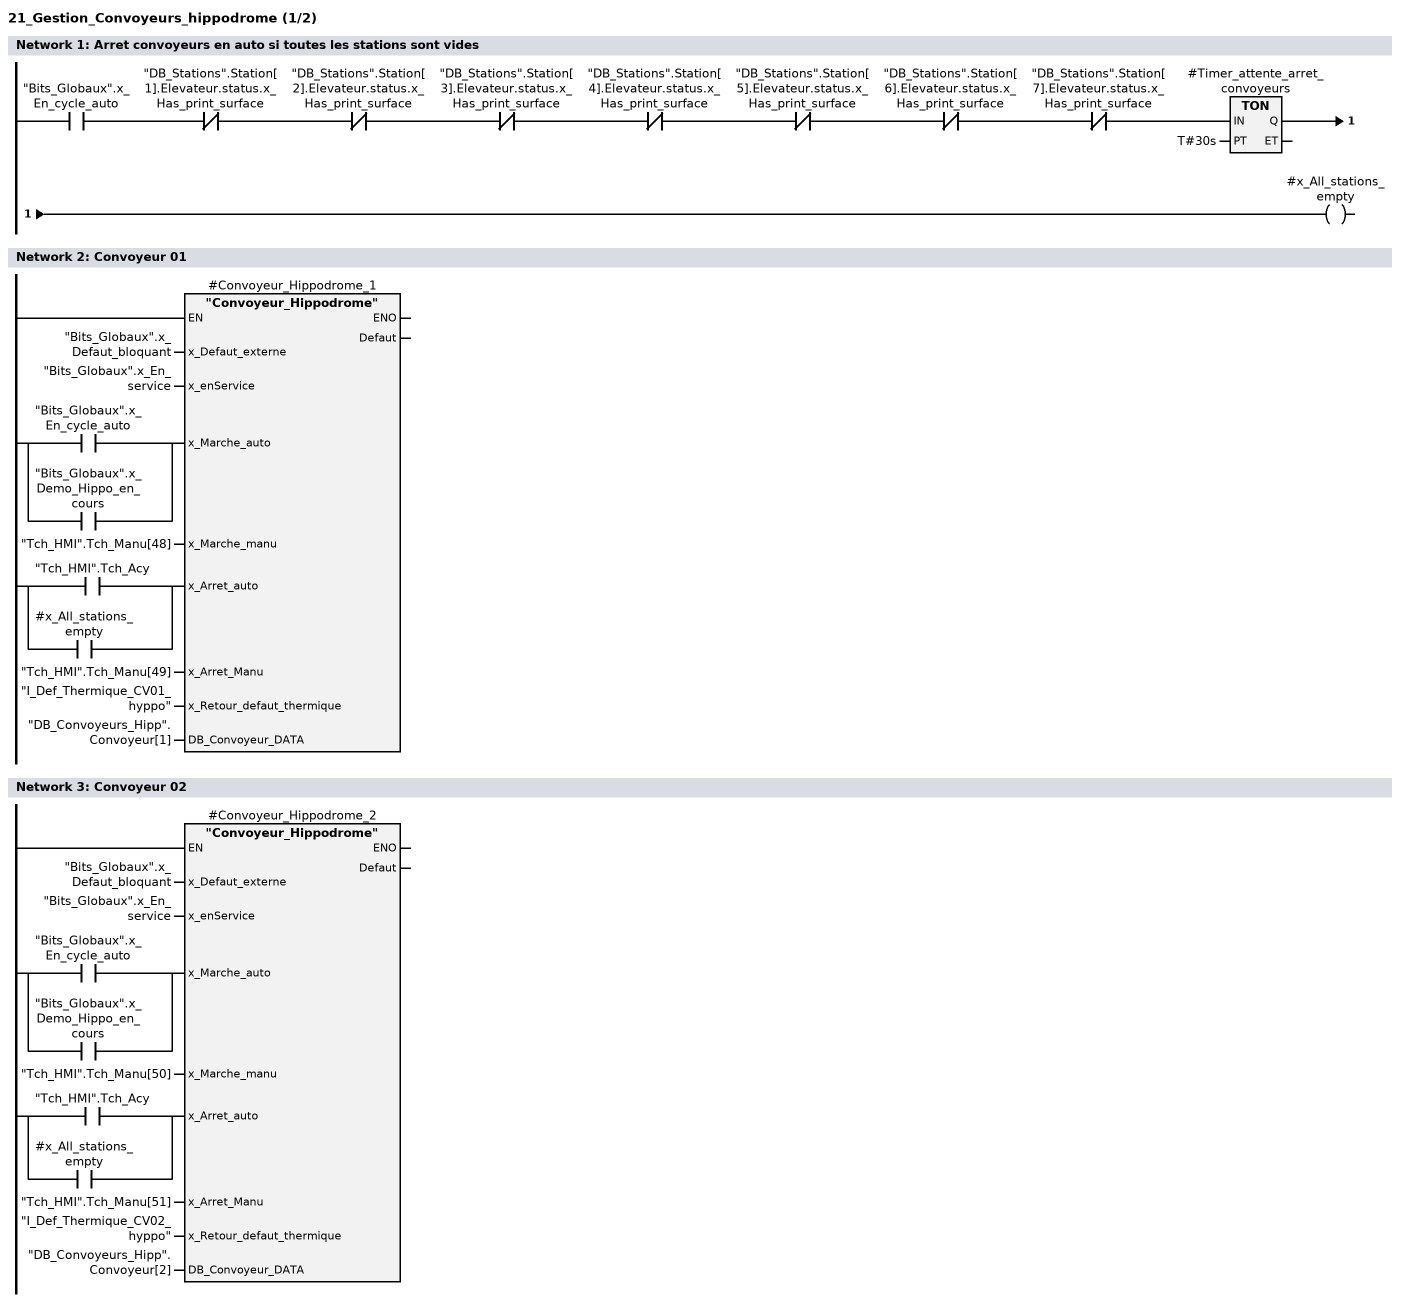
   #Timer_attente_arret_convoyeurs(IN := "Bits_Globaux".x_En_cycle_auto AND NOT "DB_Stations".Station[1].Elevateur.status.x_Has_print_surface AND NOT "DB_Stations".Station[2].Elevateur.status.x_Has_print_surface AND NOT "DB_Stations".Station[3].Elevateur.status.x_Has_print_surface AND NOT "DB_Stations".Station[4].Elevateur.status.x_Has_print_surface AND NOT "DB_Stations".Station[5].Elevateur.status.x_Has_print_surface AND NOT "DB_Stations".Station[6].Elevateur.status.x_Has_print_surface AND NOT "DB_Stations".Station[7].Elevateur.status.x_Has_print_surface,   // TON
                           PT := T#30s);
   #x_All_stations_empty := #Timer_attente_arret_convoyeurs.Q;
END_REGION

REGION Network 2: Convoyeur 01
   RUNG wire#powerrail
      #Convoyeur_Hippodrome_1(x_Marche_auto := wire#w1, x_Arret_auto := wire#w2, x_Defaut_externe := "Bits_Globaux".x_Defaut_bloquant, x_enService := "Bits_Globaux".x_En_service, x_Marche_manu := "Tch_HMI".Tch_Manu[48], x_Arret_Manu := "Tch_HMI".Tch_Manu[49], x_Retour_defaut_thermique := "I_Def_Thermique_CV01_hyppo", DB_Convoyeur_DATA := "DB_Convoyeurs_Hipp".Convoyeur[1], Defaut =>)
   END_RUNG
   RUNG wire#powerrail
      Contact( "Bits_Globaux".x_En_cycle_auto )
   END_RUNG wire#w1
   RUNG wire#powerrail
      Contact( "Bits_Globaux".x_Demo_Hippo_en_cours )
   END_RUNG wire#w1
   RUNG wire#powerrail
      Contact( "Tch_HMI".Tch_Acy )
   END_RUNG wire#w2
   RUNG wire#powerrail
      Contact( #x_All_stations_empty )
   END_RUNG wire#w2
   // the same network as SCL:
   #Convoyeur_Hippodrome_1(x_Defaut_externe := "Bits_Globaux".x_Defaut_bloquant,   // "Convoyeur_Hippodrome"
                           x_enService := "Bits_Globaux".x_En_service,
                           x_Marche_auto := "Bits_Globaux".x_En_cycle_auto OR "Bits_Globaux".x_Demo_Hippo_en_cours,
                           x_Marche_manu := "Tch_HMI".Tch_Manu[48],
                           x_Arret_auto := "Tch_HMI".Tch_Acy OR #x_All_stations_empty,
                           x_Arret_Manu := "Tch_HMI".Tch_Manu[49],
                           x_Retour_defaut_thermique := "I_Def_Thermique_CV01_hyppo",
                           DB_Convoyeur_DATA := "DB_Convoyeurs_Hipp".Convoyeur[1]);
END_REGION

